(* IEC 61131-3 sources: daoli-st-library/DL_Algo (part 15) *)

(* ---- FB_DL_InputShaperZv.st ---- *)
(*
  ==================================================================
  组件名 Component  : FB_DL_InputShaperZv
  分类   Category   : DL_Algo
  复杂度 Complexity  : 中
  版本   Version    : 1.0.1
  功能   Purpose    : ZV（Zero Vibration）双脉冲输入整形器。按阻尼比 ζ 与固有频率
                      ωn 合成两脉冲序列（幅值 1/(1+A) 与 A/(1+A)，间隔 Δt），
                      触发沿到达时先出首脉冲，经 Δt 后出次脉冲，用于抑制指令
                      阶跃激起的残余振动。
  来源   Source     : self-std（公开控制理论 ZV 整形器语义）
  溯源   Origin     : ZV 输入整形属公开控制理论（Singer & Seering 公开文献语义），
                      道莅 clean-room 自研实现，未复制任何厂商私有库源码。
  平台   Platform   : 纯 IEC 61131-3（EXPT / SQRT / TON / R_TRIG / 标准转换函数）
  分工声明 Split     : 与 FB_DL_NotchFilter（反馈侧频域抑制属主）分工——后者对
                      测量信号做在线滤波；本件只整形前馈指令时序，不接管反馈、
                      不做滤波、不判机械到位。
  作者   Author     : 道莅代码库 · PLC 编程专家（R60）
  归属 Ownership     : E_DL_ZvPhase 属主为本文件（全库唯一定义，R264）；
                      引用件只引用不重声明（D13 返修补行）。
  ------------------------------------------------------------------
  边界 Boundary     :
                      一 时间口径单一化（R342）：Δt 内部一律以秒计算，转 TIME 时
                         统一乘 1000 后经 LREAL_TO_TIME 落毫秒，禁跨日历类型链；
                      二 采样约定：首脉冲在触发沿当拍输出，次脉冲在 Δt 到期拍
                         输出，两脉冲均为单拍（统一出口段每拍先预置 FALSE，R256）；
                      三 有限性闸显式枚举全部浮点输入（R272 自证：声明区 LREAL
                         输入共 2 个——fWn 与 fZeta——闸内逐个引用，无遗漏）；
                      四 域闸：fWn ≤ 0 判故障级码并冻结输出；ζ 域 [0, 0.95) 钳位，
                         越域置信息级码（ζ = 0 为无阻尼极限，取 A = 1 双等幅脉冲，
                         √(1−ζ²) = 1 结构性安全）；
                      五 使能 bEnable = FALSE 时语义为「冻结保持 + 清未决次脉冲」
                         （不再出脉冲，幅值与间隔保持末次有效值）——R191 声明行；
                      六 故障解除路径：eFault 相由复位沿迁回空闲并清锁存（bReset
                         为输入引脚，恒可达，R152 自证）；
                      七 时序滞后声明（D12 返修登记）：tonGap 的 PT 取上拍
                         _tDelay（段 0 刷新先于段 3 参数换算），ωn 突变拍 Δt
                         生效滞后一扫描拍；上层如需同拍生效，须在触发前一拍
                         稳定参数（显式声明，非遗漏）。
  错误码   Codes    :
    16#0002_0610【信息级】阻尼比 ζ 越域已钳位到 [0, 0.95)
    16#0002_0611【故障级】浮点入参非有限（NaN / Inf），输出冻结
    16#0002_0612【故障级】固有频率 ωn ≤ 0（域非法），输出冻结
  验收   Acceptance :
    算法已证（脚本）：未跑 ｜ 编译器已证（三平台）：未跑
    V1 ωn=10 rad/s、ζ=0 → A=1、幅值各 0.5、Δt=0.314159 s（314 ms）
    V2 ωn=10 rad/s、ζ=0.3 → A=0.371、幅值 0.7290/0.2710、Δt=0.3296 s
    V3 ζ=1.5 → 钳到 0.95、码 0610、序列仍出（bValid = TRUE）
    V4 ωn=0 → 码 0612、两脉冲恒假、eState = eFault
  修订记录 Revision  :
    2026-11-21  v1.0.0  R60 首版（批 2 · 序号 8）
    2026-11-21  v1.0.1  R61 返修：D12 边界段声明 tonGap PT 一拍滞后口径；
                        D13 补 E_DL_ZvPhase 属主 Ownership 行
  ==================================================================
*)

TYPE E_DL_ZvPhase :
(
    eIdle  := 0,  // 空闲：无未决次脉冲 / idle, no pending second pulse
    eWaitB := 10, // 等次脉冲：首脉冲已出，Δt 计时中 / waiting for the second pulse while the gap runs
    eFault := 20  // 故障：参数非法，输出冻结 / fault, the parameters are illegal and the outlet is frozen
);
END_TYPE

FUNCTION_BLOCK FB_DL_InputShaperZv
VAR_INPUT
    bEnable : BOOL := TRUE;       // 使能，FALSE 时冻结保持并清未决脉冲（边界五）/ the enable, false freezes and clears the pending pulse
    bTrig   : BOOL := FALSE;      // 整形触发电平，上升沿发起双脉冲序列 / the shaping trigger, the rising edge starts the pair
    bReset  : BOOL := FALSE;      // 复位沿：清故障锁存与未决序列并回空闲 / the reset edge, clears the latch and the pending pair
    fWn     : LREAL := 10.0;      // 固有角频率 [弧度每秒]，必须 > 0 / the natural angular frequency, must be positive
    fZeta   : LREAL := 0.1;       // 阻尼比 [-]，域 [0, 0.95) / the damping ratio inside the half open domain
END_VAR
VAR_OUTPUT
    bPulseA : BOOL := FALSE;      // 首脉冲单拍（触发沿当拍）[-] / the first pulse on the trigger scan
    bPulseB : BOOL := FALSE;      // 次脉冲单拍（Δt 到期拍）[-] / the second pulse on the expiry scan
    fAmpA   : LREAL := 0.5;       // 首脉冲幅值系数 [-]，与次脉冲之和为一 / the first amplitude coefficient
    fAmpB   : LREAL := 0.5;       // 次脉冲幅值系数 [-] / the second amplitude coefficient
    tDelay  : TIME := T#0S;       // 双脉冲间隔 Δt [毫秒] / the gap between the two pulses
    eState  : E_DL_ZvPhase;       // 主状态机当前态 [状态] / the current state of the main machine
    bValid  : BOOL := FALSE;      // 参数有效且序列可用标志 [-] / the parameters valid and the pair usable flag
    bError  : BOOL := FALSE;      // 故障锁存位 [-] / the latched fault bit
    eErr    : UDINT := 16#0000_0000; // 错误码，0 = 正常 / the error code, zero is ok
END_VAR
VAR
    _bInit    : BOOL := FALSE;                       // 首拍初始化标志（R310）/ the first scan flag
    _eState   : E_DL_ZvPhase := E_DL_ZvPhase.eIdle;  // 内部状态寄存器，段 4 唯一写点 / the internal state register, single writer
    _bPulseA  : BOOL := FALSE;                       // 首脉冲内部位，段 1 预清段 6 映射 / the internal first pulse bit, preset then mapped
    _bPulseB  : BOOL := FALSE;                       // 次脉冲内部位，段 1 预清段 6 映射 / the internal second pulse bit, preset then mapped
    _bPending : BOOL := FALSE;                       // 未决次脉冲位（间隔计时使能源）/ the pending second pulse flag driving the gap timer
    _bFault   : BOOL := FALSE;                       // 故障锁存副本（仅复位沿清除）/ the fault latch copy, cleared only on the reset edge
    _bFin     : BOOL := FALSE;                       // 浮点有限性闸结果（逐拍重算）/ the finiteness gate result, recomputed every scan
    _fZetaUse : LREAL := 0.0;                        // 钳位后的阻尼比工作副本 [-] / the clamped damping ratio copy
    _fA        : LREAL := 0.0;                       // 幅值比 A = exp(−ζπ/√(1−ζ²)) [-] / the amplitude ratio
    _fRoot     : LREAL := 1.0;                       // √(1−ζ²) 工作副本 [-] / the root working copy
    _fDtSec    : LREAL := 0.0;                       // 双脉冲间隔 [秒] / the gap in seconds
    _tDelay    : TIME := T#0S;                       // 内部间隔副本，段 6 单点映射 / the internal gap copy, mapped once in segment six
    rtTrig     : R_TRIG;                            // 触发沿实例，段 0 无条件刷新 / the trigger edge instance, refreshed unconditionally
    tonGap     : TON;                               // 间隔定时器，段 0 无条件刷新 / the gap timer, refreshed unconditionally
END_VAR
VAR CONSTANT
    DL_ZV_ZETAMAX : LREAL := 0.95;                  // 阻尼比上界（开区间）[-] / the damping ratio upper bound, exclusive
    DL_ZV_PI      : LREAL := 3.14159265358979323846; // 圆周率（LREAL 精度字面量，R51）/ the pi constant at the long real precision
    DL_ZV_E       : LREAL := 2.71828182845904523536; // 自然常数（EXPT 底数，禁厂商 EXP 方言）/ the natural base used with the standard power operator
    DL_ZV_MS      : LREAL := 1000.0;                // 秒到毫秒的换算因子 [毫秒每秒] / the seconds to milliseconds factor
END_VAR

// 段 0｜沿检测与间隔定时器无条件周期刷新（禁入分支，R7；IN 串故障锁存门控，FB50-1）/ segment 0, the unconditional refresh with the latch gate
rtTrig(CLK := bTrig); // 触发沿 / the trigger edge
tonGap(IN := _bPending AND _bFin AND (NOT _bFault), PT := _tDelay); // 间隔计时：未决且参数有效且无锁存 / the gap timing only while pending and valid

// 段 1｜首拍初始化与单拍标志预清（仅单拍标志入清单，R32 FB32-1；R256）/ segment 1, the first scan init and the one shot preset
IF NOT _bInit THEN // 首拍一拍 / the first scan
    _bInit := TRUE; // 置首拍标志 / raise the first scan flag
    _bPending := FALSE; // 未决位显式清零 / clear the pending flag explicitly
    _bFault := FALSE; // 故障锁存显式清零 / clear the fault latch explicitly
    _eState := E_DL_ZvPhase.eIdle; // 状态显式落空闲 / place the state to idle explicitly
END_IF
_bPulseA := FALSE; // 首脉冲预清零 / preset the first pulse false
_bPulseB := FALSE; // 次脉冲预清零 / preset the second pulse false

// 段 2｜参数有限性闸：显式枚举全部浮点输入 fWn 与 fZeta（R272 覆盖自证，边界三）/ segment 2, the finiteness gate enumerating every floating input
_bFin := (fWn = fWn) AND ((fWn - fWn) = (fWn - fWn)) AND (fZeta = fZeta) AND ((fZeta - fZeta) = (fZeta - fZeta)); // NaN 自反判 + Inf 差值自减判，两输入逐项 / the NaN reflexive and Inf difference tests on both inputs

// 段 3｜参数域闸：频率正域与阻尼比钳位（域闸覆盖参与换算的每个引脚，边界四）/ segment 3, the domain gate covering every pin used in the computation
IF NOT _bFin THEN // 非有限参数 / a non finite parameter
    _bFault := TRUE; // 锁存故障（段 5 迁移相）/ latch the fault, the segment five migrates the phase
ELSIF fWn <= 0.0 THEN // 频率域非法 / an illegal frequency domain
    _bFault := TRUE; // 锁存故障 / latch the fault
ELSE // 参数域合法：计算整形系数 / the parameters are legal, compute the shaping coefficients
    IF fZeta < 0.0 THEN // 阻尼比低于下界 / the damping below the floor
        _fZetaUse := 0.0; // 钳到零（无阻尼极限）/ clamp to zero, the undamped limit
    ELSIF fZeta >= DL_ZV_ZETAMAX THEN // 阻尼比达上界 / the damping at the bound
        _fZetaUse := 0.84375; // 钳到域几何内点 27/32（落在 [0, 0.95) 内，二级回退，R117）/ clamp to the interior point 27 over 32
    ELSE // 域内 / inside the domain
        _fZetaUse := fZeta; // 原值接管 / take the value as is
    END_IF
    _fRoot := SQRT(1.0 - _fZetaUse * _fZetaUse); // √(1−ζ²)：ζ ≤ 0.95 保证 > 0.31（结构性安全）/ the root is provably positive
    _fA := EXPT(DL_ZV_E, 0.0 - _fZetaUse * DL_ZV_PI / _fRoot); // A = exp(−ζπ/√(1−ζ²)) / the amplitude ratio
    fAmpA := 1.0 / (1.0 + _fA); // 首脉冲幅值（除子 ≥ 1 恒正）/ the first coefficient with a divisor of at least one
    fAmpB := _fA / (1.0 + _fA); // 次脉冲幅值 / the second coefficient
    _fDtSec := DL_ZV_PI / (fWn * _fRoot); // Δt = π/(ωn√(1−ζ²)) [秒] / the gap in seconds
    _tDelay := LREAL_TO_TIME(_fDtSec * DL_ZV_MS); // 秒口径单一化后落毫秒（R342）/ the single second domain converted to milliseconds
END_IF

// 段 4｜主状态机（ENUM + CASE，ELSE 拦非法态）/ segment 4, the main machine with the illegal state guard
CASE _eState OF
    E_DL_ZvPhase.eIdle: // 空闲相：等触发沿 / the idle phase waiting for the trigger edge
        IF bEnable AND _bFin AND (NOT _bFault) AND (fWn > 0.0) AND rtTrig.Q THEN // 迁入判据带全量闸位复检（R274）/ the entry with the full gate recheck
            _bPulseA := TRUE; // 首脉冲（触发沿当拍，边界二）/ the first pulse on the trigger scan
            _bPending := TRUE; // 置未决次脉冲 / raise the pending second pulse
            _eState := E_DL_ZvPhase.eWaitB; // 迁入等次脉冲相 / enter the waiting phase
        END_IF
    E_DL_ZvPhase.eWaitB: // 等次脉冲相 / the waiting phase
        IF tonGap.Q THEN // 间隔到期：出次脉冲 / the gap expired, raise the second pulse
            _bPulseB := TRUE; // 次脉冲单拍 / the second pulse
            _bPending := FALSE; // 清未决位 / clear the pending flag
            _eState := E_DL_ZvPhase.eIdle; // 迁回空闲 / back to idle
        ELSIF (NOT bEnable) OR (NOT _bFin) OR _bFault THEN // 出口二：失能 / 参数转非有限 / 锁存（前置条件消失）/ the second exit with the prerequisite gone
            _bPending := FALSE; // 清未决位（弃用序列，不出次脉冲）/ discard the pending pair
            _eState := E_DL_ZvPhase.eIdle; // 迁回空闲 / back to idle
        END_IF
    E_DL_ZvPhase.eFault: // 故障相：锁存保持，等复位沿（解除可达，边界六）/ the fault phase held until the reset edge
        IF bReset THEN // 复位电平（复位作用域：清锁存 + 清未决 + 迁相位）/ the reset with the declared scope
            _bFault := FALSE; // 清故障锁存 / clear the fault latch
            _bPending := FALSE; // 清未决序列 / clear the pending pair
            _eState := E_DL_ZvPhase.eIdle; // 故障相迁出边回空闲 / the exit edge back to idle
        END_IF
    ELSE // 非法枚举值拦截 / the illegal enumeration guard
        _eState := E_DL_ZvPhase.eIdle; // 落回空闲 / force back to idle
        _bFault := TRUE; // 置故障锁存 / latch the fault
END_CASE

// 段 5｜故障锁存迁移闸（置于解除段之后防同拍抢迁，R258）/ segment 5, the fault latch to phase gate placed after the release
IF _bFault AND (_eState <> E_DL_ZvPhase.eFault) THEN // 已锁存但不在故障相 / latched but not in the fault phase
    _eState := E_DL_ZvPhase.eFault; // 迁入故障相 / enter the fault phase
END_IF

// 段 6｜统一出口（内部副本单点映射，R180；故障码锁存回放，R187）/ segment 6, the unified outlet
bPulseA := _bPulseA AND bEnable; // 首脉冲出口（失能不出脉冲）/ the first pulse outlet gated by the enable
bPulseB := _bPulseB AND bEnable; // 次脉冲出口（失能不出脉冲）/ the second pulse outlet gated by the enable
tDelay := _tDelay; // 间隔出口 / the gap outlet
eState := _eState; // 状态出口 / the state outlet
bError := _bFault; // 故障位出口（与锁存同源）/ the fault bit outlet from the same latch
bValid := _bFin AND (fWn > 0.0) AND (NOT _bFault); // 参数可用标志（逐拍重算）/ the usable flag recomputed every scan
IF _bFault THEN // 故障锁存回放优先 / the latched fault replays first
    IF NOT _bFin THEN // 非有限成因（独立码值，R190）/ the non finite cause with its own code
        eErr := 16#0002_0611; // 故障级：浮点入参非有限 / fault grade, a non finite floating input
    ELSE // 频率域成因 / the frequency domain cause
        eErr := 16#0002_0612; // 故障级：固有频率非正 / fault grade, the natural frequency is not positive
    END_IF
ELSIF ABS(_fZetaUse - fZeta) > 1.0E-9 THEN // 阻尼比被钳位（浮点差值比较，禁等号；信息级逐拍重算）/ the damping clamped, compared by tolerance
    eErr := 16#0002_0610; // 信息级：阻尼比越域已钳位 / informational, the damping clamped
    bError := FALSE; // 信息级不置 bError（R45 配对口径：仅故障级置位）/ the informational code never raises the fault bit
ELSE // 无事件 / no event
    eErr := 16#0000_0000; // 正常 / ok
END_IF
END_FUNCTION_BLOCK

(* ---- FB_DL_Integrator.st ---- *)
(*==============================================================================
 * 组件名称 (Component)  : FB_DL_Integrator
 * 所属子库 (Sublibrary) : DL_Algo
 * 当前版本 (Version)    : 1.0.1
 * 兼容性   (Platform)   : CODESYS 3.5 / TwinCAT 3 / 汇川 InoProShop / Machine Expert
 *                         仅依赖 Standard.library（MIN / MAX / ABS / LREAL_TO_REAL），零厂商方言
 * 功能描述 (Function)   : 梯形法离散积分器：fSum += (fIn + fInPrev)/2 · fDt，
 *                         精度高于矩形法，对缓变信号无系统偏差。内部以 LREAL
 *                         双精度累加、输出转 REAL，防长时累计的舍入漂移。
 *                         带上下限限幅（触限保持）、保持（bHold）、电平复位
 *                         （bReset）、跟踪回投（bTrack）。现场用途：流量累计
 *                         （总量表）、速度→位移、电量/电能累计。
 * 开源溯源 (Origin)     : 原创实现。双精度累加思想源自 OSCAT Basic 的
 *                         FT_INT2 误差抑制行为定义（EPL-2.0），clean-room
 *                         编写，未复制任何源码。
 * 本文件内含       : TYPE  E_DL_IntState（配套枚举，归属 DL_Algo）
 *                    FB    FB_DL_Integrator
 * 依赖     (Depends)    : 无 DL_ 内部依赖；Standard.library: LREAL_TO_REAL
 * 红线自检 (Redline)    : R1 ✓ 零全局变量表与外部变量引用 ｜ R2 ✓ 零物理 IO 地址直写
 *                         R3 ✓ 纯 IEC 61131-3 ｜ R4 ✓ 量程对调+溢出钳位+非有限值拒绝
 *                         R5 ✓ 全变量中英双语同行注释 ｜ R6 ✓ 五态 ENUM+CASE+ELSE
 *                         R7 N/A（无定时器/边沿实例）
 * 【边界披露 / Boundary disclosure】
 *   B1 rOutMin > rOutMax：自动对调并置 16#0002_0001，不中断扫描。
 *   B2 复位优先于积分：bReset 电平触发，复位拍不积分（先判 bReset）。
 *   B3 输入非有限值（NaN 或幅值超 1.0E30）：本拍拒绝积分、保持累加器、
 *      fInPrev 不同步，置 16#0002_0004。
 *   B4 累加器幅值超 1.0E30：强制钳位防 LREAL 溢出，置 16#0002_0001。
 *   B5 保持期（bHold 或未使能）不积分，fInPrev 亦不更新，恢复时无历史跳变。
 *   B6 触限后每拍仍尝试积分：输入反向或限幅放宽时自动恢复，无需复位。
 * 【验收向量 / Acceptance vectors】
 *   V1  fIn=10 EU 恒定，tSampleTime=100MS，1s 后 fOut≈10 EU·s（梯形法与
 *       解析值一致，矩形法会偏 0.5 EU·s，对比可见梯形优势）
 *   V2  fIn 由 0 线性升至 10（每拍 +1），1s 后 fOut≈5.05 EU·s（与解析积分一致）
 *   V3  rOutMax=3，V1 持续 → fOut 钳位 3、bLimitHigh=TRUE、状态 eLimited
 *   V4  bHold=TRUE → fOut 冻结；释放后从冻结值继续
 *   V5  bReset 一拍 → fOut=0、fInPrev 同步当前输入（防复位后首拍尖峰）
 *   V6  bTrack 一拍（fTrackValue=100）→ fOut=100，无扰动回投
 *   V7  fIn=NaN → 16#0002_0004，fOut 保持，累加器不动
 * 修订历史 (Revision)   :
 *   2026-11-15  v1.0.0  首版入库（Round 04 · Phase 3 · DL_Algo 批次）
 *   2026-11-15  v1.0.1  阶段五终审精修：首扫自动跟踪判据修复（原 bInit 判据
 *                       反向，bTrack 一次后累加器被永久锁死为跟踪值）
 *============================================================================*)

(*-----------------------------------------------------------------------------
 * 枚举: E_DL_IntState（归属 DL_Algo，与 FB_DL_Integrator 同文件）
 * 含义: 积分器状态机离散状态。数值步长留空位便于后续插态而不破坏已有工程。
 *----------------------------------------------------------------------------*)
TYPE E_DL_IntState :
(
    eIdle        := 0,   // 空闲态：未使能，累加器保持 / Idle state, accumulator held
    eHold        := 10,  // 保持态：操作员请求冻结累加 / Hold state, accumulation frozen on request
    eIntegrating := 20,  // 积分态：梯形法逐拍累加 / Integrating, trapezoidal accumulation
    eLimited     := 30,  // 触限态：累加器停在限幅值，反向输入自动恢复 / Limited, auto recovers on reverse input
    eFault       := 99   // 故障兜底态：非法状态拦截，自动回空闲 / Fault fallback, auto recover to idle
);
END_TYPE

(*==============================================================================
 * 功能块: FB_DL_Integrator
 * 调用约定: 每个扫描周期无条件调用一次；bReset 电平触发（保持 TRUE 即持续清零）。
 * 无状态泄漏: 全部状态驻留于实例私有 VAR，可多实例并行互不影响。
 * 精度披露: 内部 LREAL 双精度累加、每拍输出转 REAL；单位为 [EU·s]
 *           （被积量 [EU] × 时间 [s]），总表类应用注意换算口径。
 *============================================================================*)
FUNCTION_BLOCK FB_DL_Integrator
VAR_INPUT
    bEnable     : BOOL := FALSE;      // 使能标志，FALSE 保持累加器 / Enable flag, FALSE holds accumulator
    fIn         : REAL := 0.0;        // 被积量 [EU]，如流量/速度/电流 / Integrated input [EU]
    rOutMin     : REAL := 0.0;        // 积分下限 [EU·s]，大于上限时自动对调 / Integral lower limit [EU·s], swapped if greater
    rOutMax     : REAL := 1.0E12;     // 积分上限 [EU·s]，长时累计防溢出 / Integral upper limit [EU·s]
    bHold       : BOOL := FALSE;      // 保持请求，TRUE 冻结累加 / Hold request, TRUE freezes accumulation
    bReset      : BOOL := FALSE;      // 复位信号，电平触发清零 / Reset signal, level triggered clear
    bTrack      : BOOL := FALSE;      // 跟踪使能，TRUE 时累加器立即跟随 fTrackValue / Track enable, accumulator follows track value
    fTrackValue : REAL := 0.0;        // 跟踪值 [EU·s]，投切无扰动基准 / Track value [EU·s], bumpless transfer reference
    tSampleTime : TIME := T#100MS;    // 采样周期 [s]，小于 10ms 钳位为 10ms / Sample time [s], clamped to 10ms
END_VAR
VAR_OUTPUT
    fOut        : REAL;               // 积分结果 [EU·s] / Integration result [EU·s]
    bLimitHigh  : BOOL;               // 触上限标志 / Upper limit reached flag
    bLimitLow   : BOOL;               // 触下限标志 / Lower limit reached flag
    bError      : BOOL;               // 故障标志（瞬时，逐拍重算） / Fault flag, transient, recomputed every scan
    uErrorId    : UDINT;              // 故障码，0 = 无故障 / Error code, 0 = no error
END_VAR
VAR
    fSumLReal   : LREAL;              // 双精度累加器 [EU·s] / Double precision accumulator [EU·s]
    fInPrev     : REAL;               // 上一拍被积量 [EU]，梯形法端点 / Previous input [EU], trapezoid endpoint
    fDt         : REAL;               // 折算后的采样周期 [s] / Converted sample period [s]
    bInFinite   : BOOL;               // 本拍输入有限值标志 / Input finite validity flag this scan
    bInit       : BOOL;               // 首扫标志：首扫自动跟踪 / First scan flag, auto track on first scan
    eState      : E_DL_IntState;      // 主状态机当前状态 / Current state of the main state machine
END_VAR
VAR CONSTANT
    DL_INT_ABS_MAX : LREAL := 1.0E30; // 累加器幅值上限 [EU·s]，防溢出 / Accumulator magnitude limit [EU·s]
END_VAR

(*------------------------------------------------------------------------------
 * 段 1｜公共参数处理（通用约定 0-1/0-2）：周期钳位、量程对调、故障码瞬时清零
 *      Common handling: sample time clamp, limit swap, transient code reset
 *-----------------------------------------------------------------------------*)
uErrorId   := 16#0000_0000;         // 故障码逐拍重算 / Error code recomputed every scan
bError     := FALSE;                // 故障标志逐拍重算 / Fault flag recomputed every scan
bLimitHigh := FALSE;                // 触限标志逐拍重算 / Limit flags recomputed every scan
bLimitLow  := FALSE;                // 触限标志逐拍重算 / Limit flags recomputed every scan

IF tSampleTime < T#10MS THEN
    fDt      := TIME_TO_REAL(T#10MS) / 1000.0; // 非法周期钳位为 10ms / Illegal period clamped to 10ms
    uErrorId := 16#0002_0002;           // 采样周期非法已钳位 / Sample time illegal, clamped
ELSE
    fDt      := TIME_TO_REAL(tSampleTime) / 1000.0; // 周期换算为秒 [s] / Period converted to seconds [s]
END_IF

IF rOutMin > rOutMax THEN
    rOutMin   := rOutMin + rOutMax;     // 三步对调第一步：求和 / Swap step one: sum
    rOutMax   := rOutMin - rOutMax;     // 三步对调第二步：得旧下限 / Swap step two: old lower limit
    rOutMin   := rOutMin - rOutMax;     // 三步对调第三步：得旧上限 / Swap step three: old upper limit
    uErrorId  := 16#0002_0001;          // 参数越界已对调 / Limits out of order, swapped
END_IF

(*------------------------------------------------------------------------------
 * 段 2｜输入合法性与复位/跟踪（边界 B2/B3、约定 0-6）
 *      Input validity and reset/track handling
 *-----------------------------------------------------------------------------*)
bInFinite := NOT (fIn <> fIn) AND (ABS(fIn) <= 1.0E30); // NaN 判别 + 幅值防御 / NaN check plus magnitude guard

IF NOT bInFinite THEN
    uErrorId := 16#0002_0004;           // 输入非有限值已拒绝 / Non-finite input rejected
END_IF

IF bTrack OR (NOT bInit) THEN
    fSumLReal := MIN(MAX(fTrackValue, rOutMin), rOutMax); // 累加器立即跟随跟踪值并限幅 / Accumulator follows track value with limits
    IF bInFinite THEN
        fInPrev := fIn;                 // 端点同步当前输入 / Endpoint synced to current input
    END_IF
    eState := eIdle;                    // 回空闲重新评估 / Back to idle for re-evaluation
    bInit  := TRUE;                     // 首扫标志置位 / First scan flag set
END_IF

IF bReset THEN
    fSumLReal := 0.0;                   // 复位优先：累加器清零 / Reset priority: accumulator cleared
    IF bInFinite THEN
        fInPrev := fIn;                 // 端点同步当前输入，防复位后尖峰 / Endpoint synced, prevents post-reset spike
    END_IF
    eState := eIdle;                    // 复位后回空闲 / Back to idle after reset
END_IF

IF NOT bEnable THEN
    eState := eIdle;                    // 未使能：强制空闲、累加器保持 / Disabled: force idle, accumulator held
END_IF

(*------------------------------------------------------------------------------
 * 段 3｜主状态机（红线 R6）：五态 ENUM + CASE + ELSE 兜底
 *      Main state machine: five-state ENUM + CASE with mandatory ELSE fallback
 *-----------------------------------------------------------------------------*)
CASE eState OF

    eIdle:  // 空闲态：使能且输入有效且未复位未保持 → 进入积分态 / Idle: enter integrating when conditions met
        IF bEnable AND bInFinite AND (NOT bReset) AND (NOT bHold) THEN
            eState := eIntegrating;     // 进入积分态（本拍先迁移，下拍起积分）/ Enter integrating, integrate from next scan
        END_IF

    eHold:  // 保持态：释放后回积分态 / Hold: resume integrating after release
        IF bEnable AND bInFinite AND (NOT bReset) AND (NOT bHold) THEN
            eState := eIntegrating;     // 恢复积分 / Resume integration
        ELSIF NOT bEnable THEN
            eState := eIdle;            // 使能跌落回空闲 / Back to idle when disabled
        END_IF

    eIntegrating:  // 积分态：梯形法逐拍累加（边界 B3 拒绝非有限值）/ Integrating: trapezoidal accumulation
        IF NOT bEnable THEN
            eState := eIdle;            // 使能跌落回空闲 / Back to idle when disabled
        ELSIF bHold THEN
            eState := eHold;            // 保持请求 / Hold request
        ELSIF bInFinite THEN
            fSumLReal := fSumLReal + (fIn + fInPrev) / 2.0 * fDt; // 梯形法累加 [EU·s] / Trapezoidal accumulation [EU·s]
            fInPrev    := fIn;          // 端点更新 / Endpoint updated
        END_IF

    eLimited:  // 触限态：每拍仍尝试积分，反向输入或限幅放宽时自动恢复（边界 B6）/ Limited: retry every scan, auto recover
        IF NOT bEnable THEN
            eState := eIdle;            // 使能跌落回空闲 / Back to idle when disabled
        ELSIF bHold THEN
            eState := eHold;            // 保持请求 / Hold request
        ELSIF bInFinite THEN
            fSumLReal := fSumLReal + (fIn + fInPrev) / 2.0 * fDt; // 继续累加（限幅兜底）/ Keep accumulating, clamp guards
            fInPrev    := fIn;          // 端点更新 / Endpoint updated
        END_IF

    eFault:  // 故障兜底态：累加器保持，自动回空闲（无锁死）/ Fault fallback: accumulator held, recover to idle
        eState := eIdle;                // 自动恢复空闲 / Auto recover to idle

    ELSE  // 非法状态拦截：任何未定义状态一律进故障态并置码 / Illegal state interception
        eState   := eFault;             // 强制故障态 / Force fault state
        uErrorId := 16#0002_0005;       // 非法状态兜底 / Illegal state fallback
        bError   := TRUE;               // 故障标志置位 / Fault flag set

END_CASE;

(*------------------------------------------------------------------------------
 * 段 4｜溢出钳位与量程限幅、输出整形（边界 B4/B1）
 *      Overflow clamp, range limiting and output shaping
 *-----------------------------------------------------------------------------*)
IF fSumLReal > DL_INT_ABS_MAX THEN
    fSumLReal := DL_INT_ABS_MAX;        // 幅值超限钳位防溢出 / Magnitude clamped against overflow
    uErrorId  := 16#0002_0001;          // 参数越界已钳位 / Value out of range, clamped
END_IF
IF fSumLReal < -DL_INT_ABS_MAX THEN
    fSumLReal := -DL_INT_ABS_MAX;       // 负向幅值钳位 / Negative magnitude clamped
    uErrorId  := 16#0002_0001;          // 参数越界已钳位 / Value out of range, clamped
END_IF

IF fSumLReal >= rOutMax THEN
    fSumLReal   := rOutMax;             // 触上限钳位 / Clamped at upper limit
    bLimitHigh  := TRUE;                // 触上限标志 / Upper limit flag
    IF bEnable AND (NOT bHold) THEN
        eState := eLimited;             // 进入触限态 / Enter limited state
    END_IF
END_IF
IF fSumLReal <= rOutMin THEN
    fSumLReal  := rOutMin;              // 触下限钳位 / Clamped at lower limit
    bLimitLow  := TRUE;                 // 触下限标志 / Lower limit flag
    IF bEnable AND (NOT bHold) THEN
        eState := eLimited;             // 进入触限态 / Enter limited state
    END_IF
END_IF

fOut := LREAL_TO_REAL(fSumLReal);       // 双精度累加器转 REAL 输出 [EU·s] / Accumulator converted to REAL output [EU·s]
END_FUNCTION_BLOCK

(* ---- FB_DL_IterSolverRunner.st ---- *)
(* ============================================================
   DL_Algo / FB_DL_IterSolverRunner ｜ v1.0.0 ｜ 2026-11-25
   功能：多方法求根运行器（0 二分 / 1 试位 / 2 割线 / 3 Illinois / 4 Brent）
         ＋括号管理＋无解与超时出口＋迭代上限防死锁。
         纯 IEC 无函数指针，采用「求值回灌协议」：本件在 fXOut 给出待求值点，
         调用方求残差后调用方法 FeedEval(fX, fF) 回灌，主体下一拍消费并给下一点。
   边界：① 括号两端同号 → eFail、码 5（无解），不空转；② 迭代上限（0=不限，默认 100）与
         总超时（0=不限，默认 T#5S）双防死锁，各自独立码（R190 归因唯一）；超时狗武装域
         覆盖 eEvalLo / eEvalHi / eRun 三相，求值相回灌断链亦能超时退出，不永久挂死；
         ③ 回灌点与待求值点
         不匹配（|Δx|>1E-9）→ 丢弃不置错；④ 复位沿作用域：清括号/计数/回灌位/锁存/
         相位，不动 _bInit；⑤ 出口非有限即落 0（N1）；⑥ 方法内不驻留跨拍状态。
   依赖：仅 IEC 61131-3（TON/R_TRIG/ABS/MIN/MAX/LIMIT）
   溯源：DLF-B-ROOTSTEP（内部原创线）｜枚举归属：E_DL_IterRunnerPhase 唯一属主
   码位：零 16# 范式；uErrId 0 无 / 1 组态 / 2 非有限 / 3 迭代上限 / 4 超时 /
         5 括号同号 / 6 非法相位
   ============================================================ *)
TYPE E_DL_IterRunnerPhase :
(
    eIdle   := 0,    // 待机：等待启动沿 / Idle, waiting for the start edge
    eEvalLo := 10,   // 求值下界：等 f(xLo) 回灌 / Waiting for the lower bound residual
    eEvalHi := 20,   // 求值上界：等 f(xHi) 回灌 / Waiting for the upper bound residual
    eRun    := 30,   // 迭代：给试算点并消费回灌 / Iterating over trial points
    eDone   := 40,   // 完成：宽度或残差达标 / Finished within tolerance
    eFail   := 50,   // 失败：无解 / 上限 / 超时 / Failed by no root, cap or timeout
    eFault  := 90    // 故障：组态或非有限锁存 / Fault latched
);
END_TYPE

FUNCTION_BLOCK FB_DL_IterSolverRunner
VAR_INPUT
    bStart   : BOOL;   // 启动，上升沿开始一轮 [-] / Start on the rising edge
    bReset   : BOOL;   // 复位，上升沿解除失败与故障 [-] / Reset on the rising edge
    fXLo     : LREAL;  // 初始括号下界 [-] / Initial lower bracket bound
    fXHi     : LREAL;  // 初始括号上界 [-] / Initial upper bracket bound
    fTol     : LREAL;  // 宽度收敛容差，域 > 0 [-] / Convergence tolerance on the width
    nMethod  : INT;    // 方法选择 0..4 [-] / Method selector
    nIterMax : INT := 100;         // 迭代上限，0 = 不限，默认 100 次（防死锁）[次] / Iteration cap, zero means unlimited
    tTimeout : TIME := T#5S;       // 总超时，0 = 不限，默认 5s（防死锁）[ms] / Overall timeout, zero means unlimited
END_VAR
VAR_OUTPUT
    bDone    : BOOL;   // 求根完成 [-] / Root finding finished
    bError   : BOOL;   // 失败或故障 [-] / Failed or faulted
    fXOut    : LREAL;  // 当前待求值点（完成时为根候选）[-] / Point to evaluate
    fResid   : LREAL;  // 末次回灌残差 [-] / Last residual fed back
    uErrId   : UDINT;  // 事件码，0 = 无事件 [-] / Event code
    nIterOut : INT;    // 已用迭代次数 [次] / Iterations consumed
END_VAR
VAR
    rtStart  : R_TRIG;                                           // 启动沿实例，段 0 无条件刷新 / Start edge
    rtReset  : R_TRIG;                                           // 复位沿实例，段 0 无条件刷新 / Reset edge
    tonTotal : TON;                                              // 总超时狗，段 0 无条件刷新 / Overall watchdog
    _eState  : E_DL_IterRunnerPhase := E_DL_IterRunnerPhase.eIdle; // 内部相位 / Internal phase
    _bInit   : BOOL := FALSE;                                    // 首扫初始化已执行 [-] / First scan init done
    _bFed    : BOOL := FALSE;                                    // 回灌到位（协议位，方法置位）[-] / Feedback ready
    _fFedX   : LREAL := 0.0;                                     // 回灌点横坐标 [-] / Fed back abscissa
    _fFedF   : LREAL := 0.0;                                     // 回灌残差 [-] / Fed back residual
    _fA      : LREAL := 0.0;                                     // 括号下界 [-] / Lower bracket bound
    _fB      : LREAL := 0.0;                                     // 括号上界 [-] / Upper bracket bound
    _fFa     : LREAL := 0.0;                                     // 下界残差 [-] / Residual at the lower bound
    _fFb     : LREAL := 0.0;                                     // 上界残差 [-] / Residual at the upper bound
    _fXCur   : LREAL := 0.0;                                     // 当前待求值点 [-] / Current point to evaluate
    _nIter   : INT := 0;                                         // 已用迭代次数 [次] / Iterations consumed
    _bFault  : BOOL := FALSE;                                    // 故障锁存位 [-] / Latched fault bit
    _bFail   : BOOL := FALSE;                                    // 失败锁存位 [-] / Latched failure bit
    _uFault  : UDINT := 0;                                       // 事件码锁存 [-] / Latched event code
    _bCfgBad : BOOL;                                             // 组态非法当拍量 [-] / Illegal configuration flag
    _bNonFin : BOOL;                                             // 入参非有限当拍量 [-] / Non-finite argument flag
    _bTmoArm : BOOL;                                             // 总超时狗武装量（三相驻留 TRUE）[-] / Watchdog arming flag
END_VAR
VAR CONSTANT
    DL_ISR_EPS : LREAL := 1.0E-9;  // 回灌点匹配与判零容差 [-] / Feedback match and zero tolerance
    DL_ISR_C_CFG : UDINT := 1;     // 码 1：组态非法 / Code one, illegal configuration
    DL_ISR_C_FIN : UDINT := 2;     // 码 2：非有限 / Code two, non-finite value
    DL_ISR_C_ITER : UDINT := 3;    // 码 3：迭代上限 / Code three, iteration cap reached
    DL_ISR_C_TMO : UDINT := 4;     // 码 4：总超时 / Code four, overall timeout
    DL_ISR_C_SGN : UDINT := 5;     // 码 5：括号同号 / Code five, bracket lost by equal signs
    DL_ISR_C_ILL : UDINT := 6;     // 码 6：非法相位 / Code six, illegal phase fallback
END_VAR

(* 方法 NextTrial：按方法选择给下一个试算点，回退固定为括号中点（必能推进）。
   参数全部经引脚传入，不访问 FB 成员，方法内无跨拍状态（R3 方法准则）。 *)
METHOD NextTrial : LREAL
VAR_INPUT
    nSel   : INT;    // 方法选择 0..4 [-] / Method selector
    fA     : LREAL;  // 括号下界 [-] / Lower bracket bound
    fB     : LREAL;  // 括号上界 [-] / Upper bracket bound
    fFa    : LREAL;  // 下界残差 [-] / Residual at the lower bound
    fFb    : LREAL;  // 上界残差 [-] / Residual at the upper bound
    fXPrev : LREAL;  // 上一步试算点 [-] / Previous trial point
    fFxPrev : LREAL; // 上一步残差 [-] / Residual at the previous trial point
END_VAR
VAR
    _fLo  : LREAL;  // 括号小端 [-] / Smaller bracket end
    _fHi  : LREAL;  // 括号大端 [-] / Larger bracket end
    _fMid : LREAL;  // 中点 [-] / Midpoint
    _fDen : LREAL;  // 差分分母 [-] / Slope denominator
    _fX   : LREAL;  // 试算点暂存 [-] / Staged trial point
END_VAR

_fLo := MIN(fA, fB);  _fHi := MAX(fA, fB);
_fMid := _fLo + (_fHi - _fLo) / 2.0;
_fX := _fMid;                                  // 缺省回退中点
CASE nSel OF
0:  _fX := _fMid;                              // 二分
1:  _fDen := fFb - fFa;                        // 试位
    IF ABS(_fDen) > DL_ISR_EPS THEN _fX := fA - fFa * (fB - fA) / _fDen; END_IF
2:  _fDen := fFxPrev - fFa;                    // 割线（最近两点差商）
    IF ABS(_fDen) > DL_ISR_EPS THEN _fX := fXPrev - fFxPrev * (fXPrev - fA) / _fDen; END_IF
3:  _fDen := (fFb / 2.0) - fFa;                // Illinois（停滞端折半）
    IF ABS(_fDen) > DL_ISR_EPS THEN _fX := fA - fFa * (fB - fA) / _fDen; END_IF
4:  IF (ABS(fFa - fFb) > DL_ISR_EPS) AND (ABS(fFa - fFxPrev) > DL_ISR_EPS)
       AND (ABS(fFb - fFxPrev) > DL_ISR_EPS) THEN   // Brent：逆二次插值
        _fX := fA * (fFb * fFxPrev) / ((fFa - fFb) * (fFa - fFxPrev))
             + fB * (fFa * fFxPrev) / ((fFb - fFa) * (fFb - fFxPrev))
             + fXPrev * (fFa * fFb) / ((fFxPrev - fFa) * (fFxPrev - fFb));
    END_IF
ELSE
    _fX := _fMid;                              // 非法方法号：回退二分
END_CASE
IF (_fX <> _fX) OR ((_fX - _fX) <> (_fX - _fX)) THEN
    NextTrial := _fMid;                        // 非有限：回退中点
ELSE
    NextTrial := LIMIT(_fLo, _fX, _fHi);       // 夹界即 N4 出口闸
END_IF
END_METHOD

(* 方法 FeedEval：调用方回灌残差。仅接受与本拍待求值点匹配的回灌（防陈旧值污染
   括号）；不匹配静默丢弃；本方法不推进相位（推进在主体 CASE）。 *)
METHOD FeedEval : BOOL
VAR_INPUT
    fX : LREAL;  // 求值点横坐标 [-] / Abscissa the host evaluated
    fF : LREAL;  // 该点残差 [-] / Residual at that abscissa
END_VAR

FeedEval := FALSE;
IF (fX <> fX) OR (fF <> fF) THEN RETURN; END_IF
IF ABS(fX - _fXCur) > DL_ISR_EPS THEN RETURN; END_IF
_fFedX := fX;  _fFedF := fF;  _bFed := TRUE;  FeedEval := TRUE;
END_METHOD

(* 段 0：沿实例与定时器无条件每拍刷新（R7） *)
rtStart (CLK := bStart);
rtReset (CLK := bReset);
(* 超时狗武装域 = 三相驻留（eEvalLo / eEvalHi / eRun）：只守 eRun 时求值相漏回灌即永久挂死无码 *)
_bTmoArm := (_eState = E_DL_IterRunnerPhase.eEvalLo)
            OR (_eState = E_DL_IterRunnerPhase.eEvalHi)
            OR (_eState = E_DL_IterRunnerPhase.eRun);
tonTotal (IN := _bTmoArm AND (NOT _bFault) AND (tTimeout > T#0S),
          PT := tTimeout);                     // tTimeout = 0 表示不限超时

(* 段 1：单拍量预清零（锁存量与回灌位不入清单，R107） *)
_bCfgBad := FALSE;  _bNonFin := FALSE;

(* 段 2：首扫与复位沿同款初始化（清锁存 / 清括号与计数 / 迁相位，R310/R311） *)
IF (NOT _bInit) OR rtReset.Q THEN
    _bInit := TRUE;  _bFault := FALSE;  _bFail := FALSE;  _uFault := 0;
    _bFed := FALSE;  _nIter := 0;  _fA := 0.0;  _fB := 0.0;  _fXCur := 0.0;
    _eState := E_DL_IterRunnerPhase.eIdle;
END_IF

(* 段 3：组态闸与非有限闸（覆盖全部参与判据的引脚，R272） *)
IF (fTol <= 0.0) OR (nMethod < 0) OR (nMethod > 4) OR (nIterMax < 0) THEN _bCfgBad := TRUE; END_IF
IF (fXLo <> fXLo) OR (fXHi <> fXHi) OR (fTol <> fTol) THEN _bNonFin := TRUE; END_IF
(* Inf 双判（正负无穷括号 = 组态非法，禁带入括号管理）：判据与出口同源于原始入参 *)
IF ((fXLo - fXLo) <> (fXLo - fXLo)) OR ((fXHi - fXHi) <> (fXHi - fXHi))
   OR ((fTol - fTol) <> (fTol - fTol)) THEN _bNonFin := TRUE; END_IF
IF (_bCfgBad OR _bNonFin) AND (NOT (_bFault OR _bFail)) THEN
    _bFault := TRUE;  _eState := E_DL_IterRunnerPhase.eFault;
    IF _bNonFin THEN
        _uFault := DL_ISR_C_FIN;      // 非有限优先归因（值与判据同源，N1）
    ELSE
        _uFault := DL_ISR_C_CFG;      // 组态非法：容差/方法号/迭代上限
    END_IF
END_IF

(* 段 4：主状态机（七相全覆盖 + ELSE 非法相位兜底） *)
CASE _eState OF

E_DL_IterRunnerPhase.eIdle:
    IF rtStart.Q THEN
        _fA := fXLo;  _fB := fXHi;  _nIter := 0;  _bFed := FALSE;
        _fXCur := fXLo;  _eState := E_DL_IterRunnerPhase.eEvalLo;   // 先求下界残差
    END_IF

E_DL_IterRunnerPhase.eEvalLo:
    IF _bFed THEN                              // 事件：回灌到位
        _fFa := _fFedF;  _bFed := FALSE;  _fXCur := _fB;
        _eState := E_DL_IterRunnerPhase.eEvalHi;
    ELSIF tonTotal.Q THEN                      // 事件缺失：超时接管（回灌断链不再永久挂死）
        _bFail := TRUE;  _uFault := DL_ISR_C_TMO;  _eState := E_DL_IterRunnerPhase.eFail;
    ELSIF ABS(_fB - _fA) <= DL_ISR_EPS THEN    // 前置消失：括号零宽
        _bFail := TRUE;  _uFault := DL_ISR_C_SGN;  _eState := E_DL_IterRunnerPhase.eFail;
    END_IF

E_DL_IterRunnerPhase.eEvalHi:
    IF _bFed THEN
        _fFb := _fFedF;  _bFed := FALSE;
        IF (ABS(_fFa) <= DL_ISR_EPS) OR (ABS(_fFb) <= DL_ISR_EPS) THEN
            _eState := E_DL_IterRunnerPhase.eDone;          // 端点已是根
        ELSIF ((_fFa > 0.0) AND (_fFb > 0.0)) OR ((_fFa < 0.0) AND (_fFb < 0.0)) THEN
            _bFail := TRUE;  _uFault := DL_ISR_C_SGN;       // 同号：无解归因
            _eState := E_DL_IterRunnerPhase.eFail;
        ELSE
            _fXCur := NextTrial(nSel := nMethod, fA := _fA, fB := _fB, fFa := _fFa,
                                fFb := _fFb, fXPrev := _fA, fFxPrev := _fFa);
            _eState := E_DL_IterRunnerPhase.eRun;
        END_IF
    ELSIF tonTotal.Q THEN                      // 事件缺失：超时接管（上界残差回灌断链亦不再挂死）
        _bFail := TRUE;  _uFault := DL_ISR_C_TMO;  _eState := E_DL_IterRunnerPhase.eFail;
    END_IF

E_DL_IterRunnerPhase.eRun:
    IF _bFed THEN
        _bFed := FALSE;  _nIter := _nIter + 1;              // 计数唯一写入点
        IF ((_fFa > 0.0) AND (_fFedF < 0.0)) OR ((_fFa < 0.0) AND (_fFedF > 0.0)) THEN
            _fB := _fFedX;  _fFb := _fFedF;                 // 回灌点与下界异号：替上界
        ELSE
            _fA := _fFedX;  _fFa := _fFedF;
        END_IF
        IF ABS(_fFedF) <= DL_ISR_EPS THEN
            _eState := E_DL_IterRunnerPhase.eDone;          // 残差达标
        ELSIF ABS(_fB - _fA) <= fTol THEN
            _eState := E_DL_IterRunnerPhase.eDone;          // 宽度达标
        ELSIF (nIterMax > 0) AND (_nIter >= nIterMax) THEN
            _bFail := TRUE;  _uFault := DL_ISR_C_ITER;
            _eState := E_DL_IterRunnerPhase.eFail;
        ELSE
            _fXCur := NextTrial(nSel := nMethod, fA := _fA, fB := _fB, fFa := _fFa,
                                fFb := _fFb, fXPrev := _fFedX, fFxPrev := _fFedF);
        END_IF
    ELSIF tonTotal.Q THEN                      // 事件缺失：超时接管（R275 事件优先）
        _bFail := TRUE;  _uFault := DL_ISR_C_TMO;  _eState := E_DL_IterRunnerPhase.eFail;
    END_IF

E_DL_IterRunnerPhase.eDone:
    IF rtStart.Q THEN                          // 启动沿重开一轮
        _bFed := FALSE;  _nIter := 0;  _fA := fXLo;  _fB := fXHi;  _fXCur := fXLo;
        _eState := E_DL_IterRunnerPhase.eEvalLo;
    END_IF

E_DL_IterRunnerPhase.eFail:
    _bFail := TRUE;                            // 失败相驻留：码位锁存回放

E_DL_IterRunnerPhase.eFault:
    _bFault := TRUE;                           // 故障相驻留：出口保持安全值

ELSE
    _bFault := TRUE;  _uFault := DL_ISR_C_ILL;  _eState := E_DL_IterRunnerPhase.eFault;
END_CASE

(* 段 5：故障迁相闸（置于解除段之后，R274） *)
IF _bFault AND (_eState <> E_DL_IterRunnerPhase.eFault) THEN
    _eState := E_DL_IterRunnerPhase.eFault;
END_IF

(* 段 6：统一出口段（判据位与实值单点裁决，N4） *)
bDone := (_eState = E_DL_IterRunnerPhase.eDone);
bError := _bFault OR _bFail;  uErrId := _uFault;  nIterOut := _nIter;
IF (_fXCur <> _fXCur) OR ((_fXCur - _fXCur) <> (_fXCur - _fXCur)) THEN
    fXOut := 0.0;                              // 非有限兜底（N1）
ELSE
    fXOut := _fXCur;
END_IF
IF (_fFedF <> _fFedF) OR ((_fFedF - _fFedF) <> (_fFedF - _fFedF)) THEN
    fResid := 0.0;
ELSE
    fResid := _fFedF;
END_IF
END_FUNCTION_BLOCK

(* ---- FB_DL_KalmanFilter1D.st ---- *)
(*==============================================================================
 * 组件名称 (Component)  : FB_DL_KalmanFilter1D
 * 所属子库 (Sublibrary) : DL_Algo
 * 当前版本 (Version)    : 1.0.0
 * 兼容性   (Platform)   : CODESYS 3.5+ / TwinCAT 3 / 汇川 InoProShop / 施耐德 Machine Expert
 *                         仅依赖 Standard.library（TON / R_TRIG / ABS），零厂商私有库
 * 功能描述 (Function)   : 标量卡尔曼滤波。状态 _fX 与协方差 _fP，逐拍「预测 → 更新」两段：
 *                         预测 _fP := _fP + fQ（随机游走过程噪声）；更新按标量卡尔曼增益
 *                         K = _fP / (_fP + fR)，用新息 |fMeas - _fX| 修正状态并压缩协方差。
 *                         野值门限：新息绝对值超 fInnovLimit → 本拍拒收（bRejected = TRUE，
 *                         不更新状态，协方差保留预测后的增大值，使下一拍更容易接受真变化）。
 *                         协方差发散保护：_fP > fPMax 持续 tDivTime → 用当拍实测重初始化并
 *                         置信息级。失能 bEnable = FALSE → 直通 fMeas 并**冻结协方差**（不归零，
 *                         保证恢复使能时无扰）。
 * 接口     (Interface)  : 输入 fMeas 实测值、fQ 过程噪声、fR 测量噪声、fInnovLimit 新息门限、
 *                         fPMax 协方差发散上限、tDivTime 发散确认时间、bEnable 使能、bReset 复位；
 *                         输出 fOut 滤波值、fPOut 当前协方差、bRejected 本拍拒收单拍位、
 *                         bDiverged 本拍重初始化单拍位、eState / eCause / bError / nErrId。
 * 边界     (Boundary)   : ① 组态闸：fQ / fR / fInnovLimit / fPMax 任一 <= 0.0、tDivTime <= T#0S、
 *                         或任一浮点引脚为 NaN → 故障锁存（NaN 自反判为判等禁令唯一例外）；
 *                         ② 除法前判除子：_fP + fR <= DL_FLOAT_EPS 时跳过更新（不产生 Inf）；
 *                         ③ 新息与状态全走容差比较，禁 `=` / `<>` 判量值；
 *                         ④ NaN 实测 → 本拍整体拒收并置信息级，**不让 NaN 进入 _fP / _fX**
 *                         （R133 / R135：非有限值绝不写入保持槽）；
 *                         ⑤ TON 一枚 + R_TRIG 一枚段 0 无条件周期刷新；
 *                         ⑥ 故障相迁出唯一路径 = bReset 上升沿；⑦ 零全局耦合（无 GVL / 无物理地址）。
 * 输出语义 (Fallback)   : 【R191 声明】bEnable = FALSE → 输出**直通** fMeas（非冻结），协方差冻结
 *                         保持末值；eFault 相 → 输出**冻结保持**末次有效估计（不清零，避免下游
 *                         把 0 当成真测量），bError 同时为真。两分支语义互不相同，均在此显式声明。
 * 解除式   (Release)    : bReset 上升沿 ∧ 组态合法 ∧〔非发散态 ∨ 本次复位已完成协方差重装〕。
 *                         自证可满足（终审两式 1）：复位沿本身在发散态执行 _fP := fR 重装，
 *                         括内第二项即为真，故解除式不存在恒假因子。反例说明：若写成单纯
 *                         「∧ 非发散态」，故障相内 _fP 不再更新 → 该项恒假 → 故障永久不可恢复，
 *                         属 R152 恒假组合反例，故本件按括内析取式实现。
 * 码表     (Codes)      : 16#0002_03AF 故障级：卡尔曼滤波故障总码（组态非法 / 非法相位），
 *                         锁存至 bReset 上升沿，归因由 eCause 承载（R190 单件单总码）；
 *                         16#0002_04B2 信息级：非故障台账事件（野值拒收 / 发散重初始化 / 除子退化跳过）。
 *                         加码反证（R90）：三类信息事件均不改变 eCause 与 bError，且 fOut 仍为
 *                         可用值，故须留痕；三类共用一码的依据是「都只要求留痕、不要求区分动作」，
 *                         区分由 bRejected / bDiverged 两个专用布尔出口承担，无需第二个码位。
 *                         码段说明：0002 段故障子带 03xx / 信息子带 04xx，本件取 03AF / 04B2
 *                         （源码实扫该两槽为空，续接同子带已用最大值，未回填碎片孔洞）。
 * 开源溯源 (Origin)     : 道莅自研 clean-room（参考公开标量卡尔曼递推式与参数域，零代码行复制）
 * 修订历史 (Revision)   : 2026-11-19  v1.0.0  R45 首版（批次 1 · 序号 5）
 *==============================================================================*)

TYPE E_DL_Kf1State :
(
    eIdle  := 0,     // 失能待使能（直通输出） / Idle, disabled, pass-through output
    eRun   := 10,    // 滤波运行 / Filtering in run
    eFault := 90     // 故障锁存相 / Fault latched phase
);
END_TYPE

TYPE E_DL_Kf1Cause :
(
    eNone       := 0,   // 无故障成因 / No cause
    eCfgIllegal := 1,   // 组态非法（含 NaN 参数） / Illegal configuration, including NaN parameters
    ePhaseBad   := 2    // 非法相位兜底 / Illegal phase fallback
);
END_TYPE

FUNCTION_BLOCK FB_DL_KalmanFilter1D
VAR_INPUT
    fMeas       : REAL := 0.0;          // 实测值 [工程单位] / Measured value
    fQ          : REAL := 0.01;         // 过程噪声方差，域 > 0.0 [工程单位²] / Process noise variance, domain > 0.0
    fR          : REAL := 0.10;         // 测量噪声方差，域 > 0.0 [工程单位²] / Measurement noise variance, domain > 0.0
    fInnovLimit : REAL := 5.0;          // 新息门限（野值判据），域 > 0.0 [工程单位] / Innovation limit, domain > 0.0
    fPMax       : REAL := 100.0;        // 协方差发散上限，域 > 0.0 [工程单位²] / Covariance divergence limit, domain > 0.0
    tDivTime    : TIME := T#5S;         // 发散确认时间，域 > T#0S [ms] / Divergence confirm time, domain > T#0S
    bEnable     : BOOL := TRUE;         // 滤波使能，FALSE 时直通并冻结协方差 [-] / Enable, FALSE passes through and freezes covariance
    bReset      : BOOL := FALSE;        // 复位命令，上升沿清故障 [-] / Reset command, rising edge clears fault
END_VAR
VAR_OUTPUT
    fOut        : REAL;                 // 滤波输出值（故障相冻结保持末值） [工程单位] / Filtered output, frozen in fault
    fPOut       : REAL;                 // 当前协方差 [工程单位²] / Current covariance
    bRejected   : BOOL;                 // 本拍野值拒收单拍位 [-] / Single-scan outlier rejection flag
    bDiverged   : BOOL;                 // 本拍发散重初始化单拍位 [-] / Single-scan divergence reinit flag
    eState      : E_DL_Kf1State;        // 状态出口，段 6 单点映射 / State outlet
    eCause      : E_DL_Kf1Cause;        // 故障成因出口（R190 归因唯一） / Fault cause outlet
    bError      : BOOL;                 // 故障锁存标志 [-] / Fault latch flag
    nErrId      : UDINT;                // 事件码，0 = 无事件 / Event code, 0 = no event
END_VAR
VAR
    _eState     : E_DL_Kf1State := E_DL_Kf1State.eIdle;   // 内部相位（CASE 唯一写入目标） / Internal phase
    _eCause     : E_DL_Kf1Cause := E_DL_Kf1Cause.eNone;   // 故障成因锁存（锁存量） / Latched cause
    tonDiv      : TON;                  // 发散确认计时，段 0 无条件调用 / Divergence confirm timer
    rtReset     : R_TRIG;               // 复位沿实例，段 0 无条件调用 / Reset edge
    _fX         : REAL;                 // 状态估计（锁存量） [工程单位] / State estimate, latched
    _fP         : REAL;                 // 状态协方差（锁存量） [工程单位²] / State covariance, latched
    _fInnov     : REAL;                 // 本拍新息 [工程单位] / Innovation this scan
    _fK         : REAL;                 // 本拍卡尔曼增益 [-] / Kalman gain this scan
    _fDen       : REAL;                 // 更新除子 _fP + fR [工程单位²] / Update divisor _fP + fR
    _bInit      : BOOL;                 // 首次初始化完成位（锁存量） [-] / Initialized flag, latched
    _bNonFin    : BOOL;                 // 实测非有限当拍量 [-] / Non-finite measurement this scan
    _bDivCond   : BOOL;                 // 协方差超上限当拍量 [-] / Covariance above limit this scan
    _bCfgBad    : BOOL;                 // 组态非法当拍量 [-] / Illegal configuration
    _bReinit    : BOOL;                 // 本次复位已做协方差重装当拍量 [-] / Covariance re-armed by this reset
    _bFault     : BOOL;                 // 故障锁存位（锁存量） / Latched fault bit
    _uFault     : UDINT;                // 故障码锁存（锁存量） / Latched fault code
    _uInfo      : UDINT;                // 信息码，每拍重算 / Info code, recomputed each scan
END_VAR
VAR CONSTANT
    DL_FLOAT_EPS : REAL := 1.0E-6;      // 浮点判零容差（除子与判等统一口径） [工程单位²] / Float epsilon for zero tests [unit2]
END_VAR

(* —— 段 0：当拍判据派生 + 定时器与沿实例无条件周期刷新 —— *)
_bNonFin := (fMeas <> fMeas) OR ((fMeas - fMeas) <> (fMeas - fMeas));       // 实测 NaN 自反 + Inf 差值自减双判（判等禁令唯一例外） / NaN and Inf detection
_bDivCond := _fP > fPMax;                                                   // 协方差超上限当拍量 / Covariance above limit
_bCfgBad := (fQ <> fQ) OR (fR <> fR) OR (fInnovLimit <> fInnovLimit) OR (fPMax <> fPMax)   // 参数 NaN 组态闸（R151 覆盖每个引脚） / NaN config gate covering every pin
            OR (fQ <= 0.0) OR (fR <= 0.0) OR (fInnovLimit <= 0.0) OR (fPMax <= 0.0)        // 正域组态闸 / Positive-domain config gate
            OR (tDivTime <= T#0S);                                                          // 时间组态闸 / Time config gate
rtReset(CLK := bReset);                                                     // 复位沿，每拍必调（R228A） / Reset edge, called every scan
tonDiv(IN := _bDivCond AND bEnable, PT := tDivTime);                        // 发散确认计时，IN 由判据派生 / Divergence timer, IN derived from verdict

(* —— 段 1：单拍量预清零（锁存量与实例不入清单，R107） —— *)
_uInfo     := 16#0000_0000;        // 信息码每拍重算 / Info recomputed every scan
bRejected  := FALSE;               // 拒收位每拍预清，唯一分支置位（R44 单拍脉冲范式） / Reject flag preset, set in one branch only
bDiverged  := FALSE;               // 重初始化位每拍预清 / Divergence flag preset
_bReinit   := FALSE;               // 复位重装标记每拍预清 / Reset re-arm marker preset
nErrId     := 16#0000_0000;        // 事件码缺省无事件 / Event code default none
bError     := FALSE;               // 故障标志每拍预清，故障分支同拍置位（R45 配对） / Flag preset

(* —— 段 2：复位沿（含发散重装）+ 组态域闸 —— *)
IF rtReset.Q THEN                                                        // 当拍复位沿 / current-scan reset edge
    _bFault := FALSE;                                                    // 清故障锁存位（锁存量） / Clear fault latch
    _uFault := 16#0000_0000;                                             // 清故障锁存码（锁存量） / Clear latched code
    _eCause := E_DL_Kf1Cause.eNone;                                      // 清成因（锁存量） / Clear latched cause
    IF _bDivCond AND (NOT _bNonFin) THEN                                 // 发散态复位：协方差重装（解除可达性关键） / Divergent reset re-arms covariance
        _fP := fR;                                                       // 协方差按测量噪声重装 / Covariance re-armed to measurement noise
        _fX := fMeas;                                                    // 状态按当拍实测重装 / State re-armed to current measurement
        _bReinit := TRUE;                                                // 标记本次复位已完成重装 / Mark re-arm done by this reset
    END_IF
    IF _eState = E_DL_Kf1State.eFault THEN
        _eState := E_DL_Kf1State.eIdle;                                  // 故障相迁出唯一路径 / Sole exit from fault phase
    END_IF
END_IF
IF _bCfgBad THEN                                                         // 组态域闸 / Configuration gate
    _uFault := 16#0002_03AF;                                             // 故障级：卡尔曼滤波故障总码 / Fault-level: filter fault code
    _bFault := TRUE;
    bError  := TRUE;                                                     // 故障标志同拍置位（R45 配对） / Error flag set same scan
    _eCause := E_DL_Kf1Cause.eCfgIllegal;                                // 归因：组态非法 / Cause: illegal configuration
END_IF

(* —— 段 3：首次初始化（仅在无故障且实测有限时取首值） —— *)
IF (NOT _bFault) AND (NOT _bInit) AND (NOT _bNonFin) THEN
    _fX := fMeas;                                                        // 首值取实测 / First value from measurement
    _fP := fR;                                                           // 协方差取测量噪声 / Covariance from measurement noise
    _bInit := TRUE;                                                      // 初始化完成（锁存量） / Initialization done
END_IF

(* —— 段 4：预测 → 更新（仅运行态执行） —— *)
IF (NOT _bFault) AND bEnable AND _bInit AND (NOT _bNonFin) THEN
    _fP := _fP + fQ;                                                     // 预测：协方差增大 / Predict, covariance grows
    IF tonDiv.Q THEN                                                     // 发散确认到：用实测重初始化 / Divergence confirmed, reinit from measurement
        _fX := fMeas;
        _fP := fR;
        bDiverged := TRUE;                                               // 单拍位：本拍做过重初始化 / Single-scan reinit flag
        _uInfo := 16#0002_04B2;                                          // 信息级：发散重初始化留痕 / Info: divergence reinit recorded
    ELSE
        _fInnov := fMeas - _fX;                                          // 新息 / Innovation
        IF ABS(_fInnov) > fInnovLimit THEN                               // 野值门限 / Outlier gate
            bRejected := TRUE;                                           // 单拍位：本拍拒收 / Single-scan reject flag
            _uInfo := 16#0002_04B2;                                      // 信息级：野值拒收留痕 / Info: outlier rejection recorded
        ELSE
            _fDen := _fP + fR;                                           // 更新除子 / Update divisor
            IF _fDen > DL_FLOAT_EPS THEN                                 // 除零前置判 / Divide-by-zero guard
                _fK := _fP / _fDen;                                      // 卡尔曼增益 / Kalman gain
                _fX := _fX + _fK * _fInnov;                              // 状态更新 / State update
                _fP := (1.0 - _fK) * _fP;                                // 协方差压缩 / Covariance shrink
            ELSE
                _uInfo := 16#0002_04B2;                                  // 信息级：除子退化跳过 / Info: degenerate divisor skipped
            END_IF
        END_IF
    END_IF
END_IF
IF (NOT _bFault) AND bEnable AND _bNonFin THEN                           // NaN 实测：本拍拒收留痕 / NaN measurement, reject and record
    bRejected := TRUE;                                                   // 单拍位：本拍拒收 / Single-scan reject flag
    _uInfo := 16#0002_04B2;                                              // 信息级：非有限实测拒收 / Info: non-finite measurement rejected
END_IF

(* —— 段 5：故障解除式（R240 全当拍量；括内析取式自证可满足） —— *)
IF rtReset.Q AND (NOT _bCfgBad) AND ((NOT _bDivCond) OR _bReinit) THEN
    _bFault := FALSE;                                                    // 清故障锁存位（锁存量） / Clear fault latch
    _uFault := 16#0000_0000;                                             // 清故障锁存码（锁存量） / Clear latched code
    _eCause := E_DL_Kf1Cause.eNone;                                      // 清成因（锁存量） / Clear latched cause
END_IF

(* —— 段 5A：故障锁存相位迁移闸 —— *)
IF _bFault AND (_eState <> E_DL_Kf1State.eFault) THEN
    _eState := E_DL_Kf1State.eFault;                                     // 锁存即入故障相 / Latch enters fault phase
END_IF

(* —— 段 6：相位机（ENUM 全成员显式标签 + ELSE 兜底，R128） —— *)
CASE _eState OF

E_DL_Kf1State.eIdle:
    IF bEnable AND _bInit AND (NOT _bFault) THEN                         // 出口 1：使能且已初始化 / Enabled and initialized
        _eState := E_DL_Kf1State.eRun;
    ELSIF _bFault THEN                                                   // 出口 2：故障锁存 / Fault latched
        _eState := E_DL_Kf1State.eFault;
    END_IF

E_DL_Kf1State.eRun:
    IF (NOT bEnable) THEN                                                // 出口 1：失能（前置条件消失，R98） / Disabled, precondition gone
        _eState := E_DL_Kf1State.eIdle;
    ELSIF _bFault THEN                                                   // 出口 2：故障锁存 / Fault latched
        _eState := E_DL_Kf1State.eFault;
    END_IF

E_DL_Kf1State.eFault:
    ;                                                                     // 故障相：仅段 5 复位沿可迁出 / Only the reset edge leaves this phase

ELSE
    _uFault := 16#0002_03AF;                                             // 故障级：非法相位兜底（归并总码） / Illegal-phase fallback
    _bFault := TRUE;
    bError  := TRUE;
    _eCause := E_DL_Kf1Cause.ePhaseBad;                                  // 归因：非法相位 / Cause: illegal phase
    _eState := E_DL_Kf1State.eFault;

END_CASE

(* —— 段 7：出口单点映射（名实同源；锁存码回放；故障相显式钳位） —— *)
IF _bFault THEN
    fOut := _fX;                                                         // 故障相冻结保持末次有效估计（R191 声明） / Frozen hold in fault
ELSIF NOT bEnable THEN
    fOut := fMeas;                                                       // 失能相直通实测（R191 声明） / Pass-through when disabled
ELSE
    fOut := _fX;                                                         // 运行相输出状态估计 / Run-phase state estimate
END_IF
IF (fOut <> fOut) OR ((fOut - fOut) <> (fOut - fOut)) THEN                // 出口非有限复检兜底 / Output non-finite recheck
    fOut := 0.0;                                                         // 非有限即归 0，绝不外溢 / Zero out, never propagate
END_IF
fPOut := _fP;                                                            // 协方差出口（锁存量回放） / Covariance outlet
IF _bFault THEN
    nErrId := _uFault;                                                   // 故障锁存码回放 / Replay latched fault code
ELSE
    nErrId := _uInfo;                                                    // 信息码 / Info code
END_IF
bError := _bFault;                                                       // 故障标志与锁存同源（名实双出口，R191） / Flag from latch
eState := _eState;                                                       // 状态出口 / State outlet
eCause := _eCause;                                                       // 成因出口 / Cause outlet

END_FUNCTION_BLOCK

(* ---- FB_DL_LaminatorPressCtrl.st ---- *)
(*
  FB_DL_LaminatorPressCtrl  —  层压机压力-时间闭环（真空段/加压段分离双目标 + 斜坡限速）/ Laminator pressure-time closed loop
  分类 Category : DL_Algo
  码位 Code     : 16#02_3_88
  段位说明      : 86/87 格由频率/三角波发生件启用，本件启用相邻 88 格（一件一码）
  版本 Version  : 1.0.0
  来源 Source   : t2-2-lbp — ROADMAP 原记 Process 属分层误记，闭环控制律按分层判定归 Algo，本轮改判并留痕
  溯源 Origin   : clean-room 实现，层压压力曲线公开工艺语义借鉴，未复制任何源码行
                  （与 FB_DL_RollCompressForceBalance 分工：那件管力平衡，本件管压力曲线跟随）
  功能 Function : 1) 六相顺控 Idle→Evac→RampPress→Hold→Release→Done，真空段/加压段目标分离；
                  2) 加压目标经 FB_DL_RateLimiter 斜坡限速（fRampRateBarS），斜坡中段由
                  FB_DL_CascadePid 主环（压力）+ 副环（执行器阀位反馈）闭环跟随；
                  3) Hold 相按配方时长 tonHold 驻留，压力越保持窗置信息级码（不静默）；
                  4) Release 相泄压 + 缩回，常压与缩回双确认才进 Done。
  边界 Boundary : ① 真空接口契约：iVac.fPressure 为负压值，深度 = −fPressure（取正深度比较）；
                  ② iActuatorFbPct 为加压执行器阀位反馈 [0..100]%（副环 PV，未接线时副环退化跟随）；
                  ③ R228-A 达标声明：四只定时器均单相独占（IN 为单相等式），跨相迁移拍 IN 必断；
                  ④ 组态域闸覆盖全部参与换算引脚；目标越上限钳制置信息级码；
                  ⑤ R228-B 达标声明：eFault 迁出 = bReset 上升沿（段 4 承载），迁出条件
                  「rtReset.Q」为输入引脚，可满足性自证成立，逐字写于此。
  依赖 Depends  : FB_DL_CascadePid / FB_DL_RateLimiter（实例化，引脚按 registry 实名）；
                  FC_DL_Hysteresis（函数调用，bState 由本件成员持有回传）；
                  I_DL_VacuumGenerator / I_DL_Cylinder（注入，不实例化）
  码表 Error codes（本件格 02_3_88，子码步进 +0x100）:
    16#0002_0188 信息级：周期完成（Done 相）
    16#0002_0288 故障级：组态非法（目标/容差/速率/时长域非法），锁存至复位
    16#0002_0388 故障级：段超时（Evac/Ramp/Release 各相独立计时），锁存至复位
    16#0002_0488 故障级：注入件故障（真空 bFault / 气缸 bFault），锁存至复位
    16#0002_0588 故障级：状态机落 ELSE 兜底（非法相位 ID），锁存至复位
    16#0002_0688 信息级：Hold 相压力越保持窗（等待回落，不置故障）
    16#0002_0788 信息级：压力目标越组态上限，已钳制

  修订历史 Revision :
    2026-11-19  v1.0.0  R39 首版（批次 2 · 序号 6）
*)

TYPE E_DL_LamPressState :
(
    eIdle      := 0,    // 空闲：等启动指令 / Idle, waiting for start
    eEvac      := 10,   // 真空段：抽气至真空目标 / Evacuation to vacuum target
    eRampPress := 20,   // 加压段：斜坡升压 + 串级闭环跟随 / Ramp press with cascade loop
    eHold      := 30,   // 保持段：配方时长驻留 + 保持窗监视 / Recipe hold with window watch
    eRelease   := 40,   // 泄压段：放气 + 缩回双确认 / Release, blow-off and retract confirm
    eDone      := 50,   // 完成：周期落定 / Done
    eFault     := 90    // 故障：组态/超时/注入件锁定 / Fault, latched
);
END_TYPE

FUNCTION_BLOCK FB_DL_LaminatorPressCtrl
VAR_INPUT
    bStart          : BOOL := FALSE;      // 启动指令（上升沿）/ Start command
    fVacTargetKpa   : REAL := 85.0;       // 真空段目标深度 [kPa]，域 > 0 / Vacuum segment target depth
    fPressTargetBar : REAL := 1.5;        // 加压段目标压力 [bar]，域 (0, fPressMaxBar] / Press segment target
    fPressMaxBar    : REAL := 2.0;        // 加压组态上限 [bar]，域 > 0 / Press configuration ceiling
    fPressActBar    : REAL := 0.0;        // 压力变送实测 [bar]（主环 PV）/ Measured pressure, master PV
    fActuatorFbPct  : REAL := 0.0;        // 执行器阀位反馈 [%]（副环 PV）/ Actuator position feedback, slave PV
    fPressTolBar    : REAL := 0.05;       // 压力跟随容差 [bar]，域 > 0 / Pressure tracking tolerance
    fRampRateBarS   : REAL := 0.05;       // 加压斜坡速率 [bar/s]，域 > 0 / Press ramp rate
    fKpM            : REAL := 1.0;        // 主环比例增益 [1] / Master loop proportional gain
    tTiM            : TIME := T#5S;       // 主环积分时间 [s] / Master loop integral time
    fKpS            : REAL := 2.0;        // 副环比例增益 [1] / Slave loop proportional gain
    tTiS            : TIME := T#1S;       // 副环积分时间 [s] / Slave loop integral time
    tEvacDur        : TIME := T#60S;      // 真空段配方时长 [ms] / Evacuation recipe duration
    tEvacTimeout    : TIME := T#120S;     // 真空段超时 [ms]，域 > 0 / Evacuation timeout
    tPressTimeout   : TIME := T#180S;     // 加压段超时 [ms]，域 > 0 / Ramp press timeout
    tHoldDur        : TIME := T#120S;     // 保持段配方时长 [ms] / Hold recipe duration
    tReleaseTimeout : TIME := T#60S;      // 泄压段超时 [ms]，域 > 0 / Release timeout
    fAtmVacKpa      : REAL := 2.0;        // 常压确认阈值 [kPa]，域 >= 0 / Atmospheric confirmation threshold
    bReset          : BOOL := FALSE;      // 复位（eFault 迁出唯一沿）/ Reset, sole fault exit edge
END_VAR
VAR_OUTPUT
    fPressSpRamp    : REAL;               // 斜坡限速后的压力设定 [bar] / Rate-limited pressure setpoint
    fPressCmdPct    : REAL;               // 串级闭环输出 [%] / Cascade closed-loop output in percent
    nSegment        : INT;                // 当前段号 [0..3]（0=真空 1=加压 2=保持 3=泄压）/ Segment index
    bCycleDone      : BOOL;               // 周期完成 / Cycle done
    nErrId          : UDINT;              // 事件码，0 = 无事件 / Event code
    eState          : E_DL_LamPressState; // 状态出口，段尾单点映射 / State outlet
END_VAR
VAR_IN_OUT
    iVac      : I_DL_VacuumGenerator;     // 真空发生器引用（注入，不实例化）/ Vacuum generator reference
    iPressCyl : I_DL_Cylinder;            // 压合气缸引用（注入，不实例化）/ Press cylinder reference
END_VAR
VAR
    fbRate     : FB_DL_RateLimiter;       // 斜坡限速实例 / Ramp rate limiter instance
    fbPid      : FB_DL_CascadePid;        // 压力串级闭环实例 / Pressure cascade loop instance
    tonEvacTo  : TON;                     // 真空段超时（单相独占）/ Evacuation timeout, single phase
    tonPressTo : TON;                     // 加压段超时（单相独占）/ Ramp press timeout, single phase
    tonHold    : TON;                     // 保持段配方计时（单相独占，PT 接配方时长）/ Hold recipe timer, single phase
    tonRelTo   : TON;                     // 泄压段超时（单相独占）/ Release timeout, single phase
    tonWch     : TON;                     // 故障观察窗，自复位 / Fault watch window, self-resetting
    rtStart    : R_TRIG;                  // 启动上升沿 / Start rising edge
    rtReset    : R_TRIG;                  // 复位上升沿 / Reset rising edge
    _eState    : E_DL_LamPressState := E_DL_LamPressState.eIdle;  // 内部相位（CASE 唯一写入目标）/ Internal phase
    _rVacDepth : REAL;                    // 真空深度暂存 [kPa] / Vacuum depth scratch
    _rPressTgt : REAL;                    // 钳制后压力目标 [bar] / Clamped press target
    _rSpRamp   : REAL;                    // 斜坡设定中间量 [bar] / Ramped setpoint working value
    _rCmdPct   : REAL;                    // 闭环输出中间量 [%] / Closed-loop output working value
    _bVacOk    : BOOL;                    // 真空到位标志 / Vacuum reached flag
    _bPressOk  : BOOL;                    // 压力入窗标志 / Pressure in-window flag
    _uFault    : UDINT;                   // 故障码锁存 / Latched fault code
    _uInfo     : UDINT;                   // 信息码，每拍重算 / Info code
    _bFault    : BOOL;                    // 故障锁存位 / Latched fault bit
    _bCfgBad   : BOOL;                    // 组态非法聚合 / Configuration invalid aggregate
END_VAR
VAR CONSTANT
    DL_LP_WATCH_PT : TIME := T#2S;      // 故障观察窗 [ms]，自复位 / Fault watch window
    DL_LP_INF_CAP  : REAL := 1.0E15;    // 非有限值筛查幅值上限 / Non-finite screening cap
END_VAR

(* —— 段 0：定时器与边沿无条件周期刷新（R182：调用语句不得置于 IF/CASE 内） —— *)
(* Stage 0, unconditional refresh of timers and edges *)
rtStart(CLK := bStart);                                           // 启动上升沿，每拍必调
rtReset(CLK := bReset);                                           // 复位上升沿，每拍必调
tonWch(IN := (NOT tonWch.Q), PT := DL_LP_WATCH_PT);               // 观察窗自复位（表达式入参）
tonEvacTo(IN := (_eState = E_DL_LamPressState.eEvac), PT := tEvacTimeout);          // 真空段超时（单相独占）
tonPressTo(IN := (_eState = E_DL_LamPressState.eRampPress), PT := tPressTimeout);   // 加压段超时（单相独占）
tonHold(IN := (_eState = E_DL_LamPressState.eHold), PT := tHoldDur);                // 保持配方计时（单相独占，PT=配方时长）
tonRelTo(IN := (_eState = E_DL_LamPressState.eRelease), PT := tReleaseTimeout);     // 泄压段超时（单相独占）

(* —— 段 1：斜坡与串级实例无条件周期刷新（依赖件每拍必调） —— *)
(* Stage 1, dependency instances refreshed unconditionally *)
fbRate(bEnable := TRUE,                                   // 限速器恒使能，跨相平滑（斜坡连续性）
       fIn := _rPressTgt,                                 // 限速输入 = 钳制后目标
       fRateUp := MAX(fRampRateBarS, 1.0E-6),             // 上升速率（下限防零速率卡死）
       fRateDown := MAX(fRampRateBarS, 1.0E-6),           // 下降速率同源
       bTrack := (_eState <> E_DL_LamPressState.eRampPress),   // 非加压相跟踪实测压力（无扰）
       fTrackValue := fPressActBar,                       // 跟踪值 = 实测压力
       tSampleTime := T#100MS);                           // 采样周期口径与限速件默认一致
_rSpRamp := fbRate.fOut;                                  // 斜坡设定中间量
fbPid(bEnable := (_eState = E_DL_LamPressState.eRampPress) OR (_eState = E_DL_LamPressState.eHold),
      fSpMaster := _rSpRamp,                              // 主环设定 = 斜坡设定
      fPvMaster := fPressActBar,                          // 主环 PV = 压力实测
      fPvSlave := fActuatorFbPct,                         // 副环 PV = 阀位反馈
      fKpM := fKpM, tTiM := tTiM, tTdM := T#0S,           // 主环参数（微分关）
      fKpS := fKpS, tTiS := tTiS, tTdS := T#0S,           // 副环参数（微分关）
      rSpSlaveMin := 0.0, rSpSlaveMax := 100.0,           // 副设定域（阀位百分比）
      rOutMin := 0.0, rOutMax := 100.0,                   // 副环输出域
      tSampleTime := T#100MS, bReset := FALSE);           // 采样周期；PID 自身不复位（相切换靠使能门控）
_rCmdPct := fbPid.fOut;                                   // 闭环输出中间量

(* —— 段 2：单拍量预清零（锁存量 _uFault/_bFault 不入清单，R187①） —— *)
_uInfo := 16#0000_0000;             // 信息码每拍重算
bCycleDone := FALSE;                // 完成出口缺省 FALSE（Done 相单点置位）
_bCfgBad := FALSE;                  // 组态非法预清零
nErrId := 16#0000_0000;             // 事件码缺省无事件

(* —— 段 3：组态域闸（覆盖全部参与判据换算的引脚，R151） —— *)
IF (fVacTargetKpa <> fVacTargetKpa) OR (fVacTargetKpa <= 0.0) OR (ABS(fVacTargetKpa) > DL_LP_INF_CAP)
   OR (fPressActBar <> fPressActBar) OR (ABS(fPressActBar) > DL_LP_INF_CAP) THEN
    _bCfgBad := TRUE;               // 真空目标/压力实测非法
END_IF
IF (fPressMaxBar <= 0.0) OR (fPressTolBar <= 0.0) OR (fRampRateBarS <= 0.0) OR (fAtmVacKpa < 0.0) THEN
    _bCfgBad := TRUE;               // 上限/容差/速率/常压阈非法
END_IF
IF (TIME_TO_DINT(tEvacTimeout) <= 0) OR (TIME_TO_DINT(tPressTimeout) <= 0)
   OR (TIME_TO_DINT(tHoldDur) <= 0) OR (TIME_TO_DINT(tReleaseTimeout) <= 0) THEN
    _bCfgBad := TRUE;               // 各段时长/超时非法
END_IF

(* —— 段 4：eFault 迁出沿（R228-B：迁出条件 rtReset.Q 为输入引脚，恒可达） —— *)
IF rtReset.Q THEN
    _bFault := FALSE;               // 清故障锁存位
    _uFault := 16#0000_0000;
    IF _eState = E_DL_LamPressState.eFault THEN
        _eState := E_DL_LamPressState.eIdle;    // 故障相迁出：回空闲（迁出边唯一且可达）
    END_IF
END_IF

(* —— 段 5：过程量只读采集与判据 —— *)
_rVacDepth := -iVac.fPressure;                // 真空深度 = 负压反馈取反 [kPa]（接口契约：负值=真空）
_bVacOk := _rVacDepth >= fVacTargetKpa;       // 真空到位判据（每拍重算）
_bPressOk := ABS(fPressActBar - _rSpRamp) <= fPressTolBar;   // 压力入窗判据（相对斜坡设定）

(* —— 段 6：相位机（只做迁移与单发命令；出口在段 8） —— *)
CASE _eState OF

E_DL_LamPressState.eIdle:
    IF _bCfgBad AND rtStart.Q THEN
        _uFault := 16#0002_0288;            // 故障级：组态非法
        _bFault := TRUE;
        _eState := E_DL_LamPressState.eFault;
    ELSIF rtStart.Q AND (NOT _bCfgBad) THEN
        IF fPressTargetBar > fPressMaxBar THEN
            _rPressTgt := fPressMaxBar;     // 压力目标越上限钳制
            _uInfo := 16#0002_0788;         // 信息级：已钳制
        ELSE
            _rPressTgt := fPressTargetBar;  // 域内直通
        END_IF
        iVac.CmdEvacuate();                 // 单发抽气指令
        _eState := E_DL_LamPressState.eEvac;    // 进真空段
    END_IF

E_DL_LamPressState.eEvac:
    IF (iVac.bFault OR iPressCyl.bFault) THEN
        _uFault := 16#0002_0488;            // 故障级：注入件故障
        _bFault := TRUE;
        iVac.CmdStop();                     // 安全侧全停
        _eState := E_DL_LamPressState.eFault;
    ELSIF tonEvacTo.Q THEN
        _uFault := 16#0002_0388;            // 故障级：真空段超时
        _bFault := TRUE;
        iVac.CmdStop();
        _eState := E_DL_LamPressState.eFault;
    ELSIF _bVacOk AND tonWch.Q THEN
        _eState := E_DL_LamPressState.eRampPress;   // 真空到位（含观察窗防抖）：进加压段
    END_IF

E_DL_LamPressState.eRampPress:
    IF (iVac.bFault OR iPressCyl.bFault) THEN
        _uFault := 16#0002_0488;
        _bFault := TRUE;
        iPressCyl.CmdStop();                // 安全侧停缸
        _eState := E_DL_LamPressState.eFault;
    ELSIF tonPressTo.Q THEN
        _uFault := 16#0002_0388;            // 故障级：加压段超时
        _bFault := TRUE;
        iPressCyl.CmdStop();
        _eState := E_DL_LamPressState.eFault;
    ELSE
        IF NOT iPressCyl.bExtended THEN
            iPressCyl.CmdExtend();          // 未到位则持续请求伸出（缸件内单发化去重）
        END_IF
        IF _bPressOk AND iPressCyl.bExtended THEN
            _eState := E_DL_LamPressState.eHold;    // 压力入窗且到位：进保持段
        END_IF
    END_IF

E_DL_LamPressState.eHold:
    IF (iVac.bFault OR iPressCyl.bFault) THEN
        _uFault := 16#0002_0488;
        _bFault := TRUE;
        iPressCyl.CmdStop();
        _eState := E_DL_LamPressState.eFault;
    ELSIF NOT _bPressOk THEN
        _uInfo := 16#0002_0688;             // 信息级：保持窗越限（等待回落，不置故障）
    ELSIF tonHold.Q THEN
        iVac.CmdBlowOff();                  // 单发放气（保持到点）
        iPressCyl.CmdRetract();             // 单发缩回
        _eState := E_DL_LamPressState.eRelease;     // 进泄压段
    END_IF

E_DL_LamPressState.eRelease:
    IF (iVac.bFault OR iPressCyl.bFault) THEN
        _uFault := 16#0002_0488;
        _bFault := TRUE;
        iPressCyl.CmdStop();
        _eState := E_DL_LamPressState.eFault;
    ELSIF tonRelTo.Q THEN
        _uFault := 16#0002_0388;            // 故障级：泄压段超时
        _bFault := TRUE;
        _eState := E_DL_LamPressState.eFault;
    ELSIF (_rVacDepth <= fAtmVacKpa) AND (NOT iPressCyl.bExtended) THEN
        _eState := E_DL_LamPressState.eDone;    // 常压 + 缩回双确认：进完成相
    END_IF

E_DL_LamPressState.eDone:
    bCycleDone := TRUE;                     // 完成出口（Done 相每拍重申）
    _uInfo := 16#0002_0188;                 // 信息级：周期完成
    IF NOT bStart THEN
        _eState := E_DL_LamPressState.eIdle;    // 指令撤销：回空闲
    END_IF

E_DL_LamPressState.eFault:
    ;                                       // 故障相：等复位沿（段 4 承载迁出）

ELSE
    _uFault := 16#0002_0588;                // 故障级：非法相位 ID 兜底
    _bFault := TRUE;
    _eState := E_DL_LamPressState.eFault;   // 强制回故障相

END_CASE

(* —— 段 7：出口单点映射（名实同源；锁存码回放，禁同拍抹除） —— *)
IF _eState = E_DL_LamPressState.eEvac THEN
    nSegment := 0;                          // 段号 0：真空
ELSIF _eState = E_DL_LamPressState.eRampPress THEN
    nSegment := 1;                          // 段号 1：加压
ELSIF _eState = E_DL_LamPressState.eHold THEN
    nSegment := 2;                          // 段号 2：保持
ELSIF _eState = E_DL_LamPressState.eRelease THEN
    nSegment := 3;                          // 段号 3：泄压
ELSE
    nSegment := -1;                         // Idle/Done/Fault：无有效段号
END_IF
fPressSpRamp := _rSpRamp;                   // 斜坡设定镜像
fPressCmdPct := _rCmdPct;                   // 闭环输出镜像
IF _bFault THEN
    nErrId := _uFault;                      // 故障锁存码回放（不在故障相按当下输入重推）
    bCycleDone := FALSE;                    // 故障相完成出口强制 FALSE（安全侧）
ELSE
    nErrId := _uInfo;                       // 信息码
END_IF
eState := _eState;                          // 状态出口单点映射

END_FUNCTION_BLOCK

(* ---- FB_DL_LeadLagCompensator.st ---- *)
(*
    FB_DL_LeadLagCompensator —— 一阶超前滞后相位校正器
    ------------------------------------------------------------------
    分类      : DL_Algo / ControlLaw
    前缀      : FB_DL_
    版本      : 1.0.0
    溯源      : 超前滞后校正 Kc·(1 + T_lead·s)/(1 + T_lag·s) 为公开经典控制判据（公共知识）；
                Tustin 双线性离散化、在线改参保状态、旁路与保持判决、错误分级与码位
                100% 自有；只借「控制器归算法层且各律独立成块」的分类组织，不复制任何
                实现代码；clean-room 重写，未复制任何闭源厂商源码，参考实现仅限 MIT/Apache 许可
    平台      : 纯 IEC 61131-3，CODESYS V3.5+ / TwinCAT 3 / InoProShop 通用
    作者      : 道莅代码库 · PLC编程专家（R19）
    ------------------------------------------------------------------
    功能说明  : 回路振荡但相位裕度不足时给前向通道加相位超前；抑制低频扰动时加滞后。
                离散化用 Tustin：a0 = 2·T_lag/Ts + 1，b0 = Kc·(1 + 2·T_lead/Ts)/a0，
                b1 = Kc·(1 − 2·T_lead/Ts)/a0，a1 = (1 − 2·T_lag/Ts)/a0。
                核心防御：① 采样周期越域或滞后时间小于采样周期，离散化极点会出单位圆，
                   此时故障级 2910 并旁路（宁可直通，不可输出病态波形）；
                ② 归一化分母 a0 前置防零判据，绝不裸除；
                ③ 增益非有限或近零即故障级 2911 并旁路——增益 0 会把回路静默掐死，
                   比报错更危险；
                ④ 输入非有限时输出保持末次有效且不旁路（旁路会把毒值直接注入执行器）；
                ⑤ 在线改参逐项比对并重算系数，历史状态保留不清零，切换无扰；
                ⑥ 输出双侧限幅，超限置 bSaturated。
                职责边界：前馈归 FeedforwardComp，纯滞后补偿归 SmithPredictor，各类滤波另件。
    错误码    : 16#0002_2901 时间常数超域已钳位 / 在线改参已重算系数（状态保留）/ 输出限幅生效——信息级，正常防御
                16#0002_2902 预留禁用（信息级，不得挪用）
                16#0002_2910 采样周期或滞后时间非法（离散化失效），旁路输出——故障级，fOut = fIn
                16#0002_2911 增益非有限或近零、输入非有限——故障级，输出保持末次有效
                16#0002_2912 预留禁用（故障级，不得挪用）
    码位总账  : 16#0002_2901 用 / 16#0002_2902 预留 ｜ 16#0002_2910 用 / 16#0002_2911 用 / 16#0002_2912 预留
    状态机    : R6 标注 N/A —— 本组件为纯函数无顺序状态机，无 CASE 可写，非法状态不可能出现
                （旁路/正常由单比特判决在段内直接给出，不存在顺序态）
    采样约定  : fbTrigReset 在本体首部无条件刷新；差分式为直接 I 型（fX1 / fY1 两状态量），
                与直接 II 型转置（单状态量）数学等价，选 I 型以保留输入输出历史供 HMI
                与改参连续性观测；时间基准全部来自 tSampleTime 引脚。
    修订记录  : 2026-11-16 v1.0.0 首次入库（R19）
*)
FUNCTION_BLOCK FB_DL_LeadLagCompensator
VAR_INPUT
    bEnable         : BOOL;                   // 使能，FALSE 旁路（输出 = 输入）/ enable, FALSE bypasses the block, output equals input
    bReset          : BOOL;                   // 复位，上升沿清内部状态 / reset, rising edge clears the internal state
    fIn             : REAL := 0.0;            // 输入（一般接偏差）[用户单位] / input, usually the control error [user unit]
    fGain           : REAL := 1.0;            // 静态增益 Kc [无量纲]，范围 -1000.0~1000.0，禁 0 / static gain [dimensionless], range -1000.0~1000.0, zero forbidden
    tLeadTime       : TIME := T#100MS;        // 超前时间常数 [ms]，范围 0~60000 / lead time constant [ms], range 0~60000
    tLagTime        : TIME := T#1S;           // 滞后时间常数 [ms]，范围 1~600000，必须 ≥ 采样周期 / lag time constant [ms], range 1~600000, must be >= the sample time
    tSampleTime     : TIME := T#100MS;        // 采样周期 [ms]，范围 1~10000 / sample time [ms], range 1~10000
    fOutLimit       : REAL := 1.0E6;          // 输出幅值限幅 [用户单位]，必须 > 0 / output magnitude limit [user unit], must be > 0
END_VAR
VAR_OUTPUT
    fOut            : REAL;                   // 校正后输出 [用户单位] / compensated output [user unit]
    bBypass         : BOOL;                   // 旁路中（参数非法或未使能）/ bypassed, illegal parameters or disabled
    bSaturated      : BOOL;                   // 输出被限幅 / output clamped
    uCoeffRev       : UDINT;                   // 系数重算次数（在线改参监视）[次] / coefficient recompute count [times]
    eErr            : UDINT;                  // 错误码，0=正常 / error id, 0=ok
    bError          : BOOL;                   // 故障标志，eErr 为故障级时 TRUE / error flag, TRUE on fault-level eErr
END_VAR
VAR
    fbTrigReset     : R_TRIG;                 // 复位上升沿实例，本体首部无条件刷新 / reset edge instance, refreshed unconditionally
    fB0             : REAL;                   // Tustin 归一化前向零次系数 [无量纲] / normalised feedforward zero-order coefficient
    fB1             : REAL;                   // Tustin 归一化前向一次系数 [无量纲] / normalised feedforward first-order coefficient
    fA1             : REAL;                   // Tustin 归一化反馈一次系数 [无量纲] / normalised feedback first-order coefficient
    fA0             : REAL;                   // Tustin 归一化分母（防零判据对象）[无量纲] / normalisation denominator, the zero guard target
    fX1             : REAL;                   // 上一拍输入历史 [用户单位] / previous input history [user unit]
    fY1             : REAL;                   // 上一拍输出历史 [用户单位] / previous output history [user unit]
    fPrevK          : REAL;                   // 上一拍增益，改参检测用 [无量纲] / previous gain for change detection [dimensionless]
    fPrevTl         : REAL;                   // 上一拍超前时间，改参检测用 [s] / previous lead time for change detection [s]
    fPrevTg         : REAL;                   // 上一拍滞后时间，改参检测用 [s] / previous lag time for change detection [s]
    fPrevTs         : REAL;                   // 上一拍采样周期，改参检测用 [s] / previous sample time for change detection [s]
    tLeadSec        : REAL;                   // 超前时间常数的秒值 [s] / lead time constant in seconds [s]
    tLagSec         : REAL;                   // 滞后时间常数的秒值 [s] / lag time constant in seconds [s]
    tTsSec          : REAL;                   // 采样周期的秒值 [s] / sample time in seconds [s]
    fLeadEff        : REAL;                   // 钳位后的超前时间 [s] / clamped lead time [s]
    fLagEff         : REAL;                   // 钳位后的滞后时间 [s] / clamped lag time [s]
    fLimitEff       : REAL;                   // 钳位后的输出限幅 [用户单位] / clamped output limit [user unit]
    bParamChg       : BOOL;                   // 在线改参标志 / parameter change flag
    bInit           : BOOL := FALSE;          // 首扫标志，初值 FALSE，判据 NOT bInit / first-scan flag, initial FALSE, tested with NOT
    nDtMs           : DINT;                   // 采样周期毫秒整数 [ms] / sample time in integer milliseconds [ms]
END_VAR
VAR CONSTANT
    DL_LL_LEAD_MAX   : TIME := T#60S;         // 超前时间上限 [ms] / lead time upper bound [ms]
    DL_LL_LAG_MAX    : TIME := T#600S;        // 滞后时间上限 [ms] / lag time upper bound [ms]
    DL_LL_GAIN_MAX   : REAL := 1000.0;        // 增益绝对值上限 [无量纲] / gain magnitude upper bound [dimensionless]
    DL_LL_DT_MAX     : TIME := T#10S;         // 采样周期上限 [ms] / sample time upper bound [ms]
    DL_LL_DT_MIN     : TIME := T#1MS;         // 采样周期下限 [ms] / sample time lower bound [ms]
    DL_FLOAT_EPS     : REAL := 1.0E-6;        // 浮点判等容差 [无量纲] / float equality tolerance [dimensionless]
    DL_LL_MICRO      : REAL := 1.0E-6;        // 微秒级容差，离散系数判定用 [无量纲] / micro tolerance for the discrete coefficients
    DL_LL_MS_PER_S   : REAL := 1000.0;        // 毫秒到秒换算因子 [ms/s] / milliseconds per second [ms/s]
    DL_LL_TWO        : REAL := 2.0;           // Tustin 分子常数 2 [无量纲] / Tustin numerator constant two [dimensionless]
    DL_LL_INF_GUARD  : REAL := 1.0E38;        // 非有限幅值判定阈值 [无量纲] / non-finite magnitude guard [dimensionless]
    DL_LL_ONE        : REAL := 1.0;           // 一值常量，归一化式用 [无量纲] / one constant used by the normalisation [dimensionless]
    DL_LL_CNT_MAX    : UDINT := 16#FFFF_FFFE; // 重算计数饱和值 [次] / recompute counter saturation value [times]
    DL_LL_ZERO       : REAL := 0.0;           // 零值常量，避免裸字面量 [无量纲] / zero constant, avoids a bare literal [dimensionless]
END_VAR

// 段 1｜边沿实例无条件周期刷新（红线：严禁放入条件分支）/ segment 1, unconditional edge refresh
fbTrigReset(CLK := bReset);

// 段 2｜输出与状态预置 / segment 2, preset outputs and status
eErr := 0;                                    // 预置无错误 / preset no error
bError := FALSE;                              // 预置无故障 / preset no fault
bBypass := FALSE;                             // 预置非旁路 / preset not bypassed
bSaturated := FALSE;                          // 预置未饱和 / preset not saturated

// 段 3｜首扫初始化（唯一合法范式：初值 FALSE，判据 NOT bInit）/ segment 3, first-scan initialisation
IF NOT bInit THEN
    fX1 := DL_LL_ZERO;                        // 输入历史清零 / clear the input history
    fY1 := DL_LL_ZERO;                        // 输出历史清零 / clear the output history
    fPrevK := DL_LL_GAIN_MAX;                 // 上一拍增益置哨兵值，首拍必触发重算 / sentinel forces a recompute on the first scan
    fPrevTl := -DL_LL_TWO;                    // 相同哨兵策略 / same sentinel strategy
    fPrevTg := -DL_LL_TWO;                    // 相同哨兵策略 / same sentinel strategy
    fPrevTs := -DL_LL_TWO;                    // 相同哨兵策略 / same sentinel strategy
    bInit := TRUE;                            // 首扫只做一次 / first scan runs once only
END_IF

// 段 4｜使能闸：未使能直接旁路 / segment 4, enable gate bypasses the block
IF NOT bEnable THEN
    bBypass := TRUE;                          // 标记旁路 / flag the bypass
    fOut := fIn;                              // 旁路即直通 / bypass means straight through
    RETURN;                                   // 失能即出口 / disabled is the exit
END_IF

// 段 5｜采样周期与滞后时间闸（离散化失效时宁可直通）/ segment 5, discretisation validity gate
IF (tSampleTime < DL_LL_DT_MIN) OR (tSampleTime > DL_LL_DT_MAX) THEN
    eErr := 16#0002_2910;                     // 采样周期非法故障码 / illegal sample time fault id
    bError := TRUE;                           // 置故障标志 / raise the error flag
    bBypass := TRUE;                          // 旁路输出 / bypass the output
    fOut := fIn;                              // 直通，不输出病态波形 / straight through, never emit a pathological waveform
    RETURN;                                   // 故障级提前返回 / early return on fault
END_IF
IF tLagTime < tSampleTime THEN
    eErr := 16#0002_2910;                     // 滞后时间小于采样周期，极点会出单位圆 / a lag shorter than the sample time pushes the pole outside the unit circle
    bError := TRUE;                           // 置故障标志 / raise the error flag
    bBypass := TRUE;                          // 旁路输出 / bypass the output
    fOut := fIn;                              // 直通 / straight through
    RETURN;                                   // 故障级提前返回 / early return on fault
END_IF

// 段 6｜增益闸（增益 0 会把回路静默掐死，必须报错并旁路）/ segment 6, gain gate
IF (fGain <> fGain) OR (fGain > DL_LL_INF_GUARD) OR (fGain < -DL_LL_INF_GUARD)
   OR (ABS(fGain) <= DL_FLOAT_EPS) OR (ABS(fGain) > DL_LL_GAIN_MAX) THEN
    eErr := 16#0002_2911;                     // 增益非法故障码 / illegal gain fault id
    bError := TRUE;                           // 置故障标志 / raise the error flag
    bBypass := TRUE;                          // 旁路输出 / bypass the output
    fOut := fIn;                              // 直通 / straight through
    RETURN;                                   // 故障级提前返回 / early return on fault
END_IF

// 段 7｜时间常数域钳位（超上限只钳位并留信息码）/ segment 7, time constant domain clamp
fLeadEff := DINT_TO_REAL(TIME_TO_DINT(tLeadTime)) / DL_LL_MS_PER_S; // 超前时间换算为秒 [s] / lead time in seconds [s]
fLagEff := DINT_TO_REAL(TIME_TO_DINT(tLagTime)) / DL_LL_MS_PER_S;   // 滞后时间换算为秒 [s] / lag time in seconds [s]
nDtMs := TIME_TO_DINT(tSampleTime);           // 采样周期取整数毫秒 [ms] / sample time in integer milliseconds [ms]
tTsSec := DINT_TO_REAL(nDtMs) / DL_LL_MS_PER_S; // 采样周期换算为秒，除子为常量 [s] / sample time in seconds, divisor is a constant [s]
IF fLeadEff < DL_LL_ZERO THEN
    fLeadEff := DL_LL_ZERO;                   // 超前时间为负无物理意义 / a negative lead time has no physical meaning
    eErr := 16#0002_2901;                     // 信息级：已钳位 / info level, clamped
END_IF
IF fLeadEff > (DINT_TO_REAL(TIME_TO_DINT(DL_LL_LEAD_MAX)) / DL_LL_MS_PER_S) THEN
    fLeadEff := DINT_TO_REAL(TIME_TO_DINT(DL_LL_LEAD_MAX)) / DL_LL_MS_PER_S; // 超前时间超上限钳位 [s] / clamp the lead time at its upper bound [s]
    eErr := 16#0002_2901;                     // 信息级：已钳位 / info level, clamped
END_IF
IF fLagEff > (DINT_TO_REAL(TIME_TO_DINT(DL_LL_LAG_MAX)) / DL_LL_MS_PER_S) THEN
    fLagEff := DINT_TO_REAL(TIME_TO_DINT(DL_LL_LAG_MAX)) / DL_LL_MS_PER_S; // 滞后时间超上限钳位 [s] / clamp the lag time at its upper bound [s]
    eErr := 16#0002_2901;                     // 信息级：已钳位 / info level, clamped
END_IF
tLeadSec := fLeadEff;                         // 记录生效超前时间 [s] / record the effective lead time [s]
tLagSec := fLagEff;                           // 记录生效滞后时间 [s] / record the effective lag time [s]

// 段 8｜输出限幅参数域钳位（0 或负值会让输出恒 0）/ segment 8, output limit clamp
fLimitEff := fOutLimit;                       // 取入参副本 / copy the input
IF (fLimitEff <> fLimitEff) OR (fLimitEff < DL_FLOAT_EPS) THEN
    fLimitEff := DL_LL_GAIN_MAX;              // 非法限幅退回常量上限 / fall back to the constant bound
    eErr := 16#0002_2901;                     // 信息级：限幅参数已收敛 / info level, the limit was converged
END_IF

// 段 9｜在线改参检测（逐项比对，命中即重算系数并保留历史状态）/ segment 9, online parameter change detection
bParamChg := (ABS(fGain - fPrevK) > DL_FLOAT_EPS)
          OR (ABS(tLeadSec - fPrevTl) > DL_FLOAT_EPS)
          OR (ABS(tLagSec - fPrevTg) > DL_FLOAT_EPS)
          OR (ABS(tTsSec - fPrevTs) > DL_FLOAT_EPS); // 改参判定 / parameter change detection
IF bParamChg THEN
    fA0 := DL_LL_TWO * tLagSec / tTsSec + DL_LL_ONE; // 归一化分母 a0 = 2·T_lag/Ts + 1 / normalisation denominator
    IF ABS(fA0) <= DL_LL_MICRO THEN
        eErr := 16#0002_2910;                 // 分母近零，离散化不可用（前置防零）/ the denominator is near zero, the discretisation is unusable
        bError := TRUE;                       // 置故障标志 / raise the error flag
        bBypass := TRUE;                      // 旁路输出 / bypass the output
        fOut := fIn;                          // 直通 / straight through
        RETURN;                               // 故障级提前返回，绝不裸除 / early return, never divide blindly
    END_IF
    fB0 := fGain * (DL_LL_TWO * tLeadSec / tTsSec + DL_LL_ONE) / fA0; // 前向零次系数 / feedforward zero-order coefficient
    fB1 := fGain * (DL_LL_ONE - DL_LL_TWO * tLeadSec / tTsSec) / fA0; // 前向一次系数 / feedforward first-order coefficient
    fA1 := (DL_LL_ONE - DL_LL_TWO * tLagSec / tTsSec) / fA0;          // 反馈一次系数 / feedback first-order coefficient
    fPrevK := fGain;                          // 记录本拍增益 / remember the gain
    fPrevTl := tLeadSec;                      // 记录本拍超前时间 / remember the lead time
    fPrevTg := tLagSec;                       // 记录本拍滞后时间 / remember the lag time
    fPrevTs := tTsSec;                        // 记录本拍采样周期 / remember the sample time
    IF uCoeffRev < DL_LL_CNT_MAX THEN
        uCoeffRev := uCoeffRev + 1;           // 重算次数饱和加一 / saturating recompute counter
    END_IF
    IF eErr = 0 THEN
        eErr := 16#0002_2901;                 // 信息级：在线改参已重算系数，状态保留 / info level, coefficients recomputed, state kept
    END_IF
    // 历史状态 fX1 / fY1 不清零：改参瞬间无扰，避免输出台阶冲击执行器 / the history is deliberately kept, so a parameter change causes no step
END_IF

// 段 10｜输入非有限闸：输出保持末次有效，且不旁路（旁路会把毒值注入执行器）/ segment 10, non-finite input gate
IF (fIn <> fIn) OR (fIn > DL_LL_INF_GUARD) OR (fIn < -DL_LL_INF_GUARD) THEN
    eErr := 16#0002_2911;                     // 输入非有限故障码 / non-finite input fault id
    bError := TRUE;                           // 置故障标志 / raise the error flag
    RETURN;                                   // 保持末次 fOut，绝不直通 / hold the last output, never pass the poison value through
END_IF

// 段 11｜复位沿清内部状态（在运算之前生效）/ segment 11, reset clears the internal state
IF fbTrigReset.Q THEN
    fX1 := DL_LL_ZERO;                        // 清输入历史 / clear the input history
    fY1 := DL_LL_ZERO;                        // 清输出历史 / clear the output history
END_IF

// 段 12｜直接 I 型差分式（两状态量，系数已归一化）/ segment 12, direct form I difference equation
fOut := fB0 * fIn + fB1 * fX1 - fA1 * fY1;    // y = b0·x + b1·x1 − a1·y1 [用户单位] / the difference equation [user unit]

// 段 13｜结果非有限复检（此时 fY1 仍是上一拍有效输出，可安全回退）/ segment 13, non-finite recheck before the state shift
IF (fOut <> fOut) OR (fOut > DL_LL_INF_GUARD) OR (fOut < -DL_LL_INF_GUARD) THEN
    eErr := 16#0002_2911;                     // 结果非有限，按输入故障同码处理 / a non-finite result shares the input fault id
    bError := TRUE;                           // 置故障标志 / raise the error flag
    fOut := fY1;                              // 回退到上一拍有效输出（位移尚未发生）/ fall back to the previous valid output, the shift has not happened yet
    RETURN;                                   // 出口 / exit
END_IF
IF fOut > fLimitEff THEN
    fOut := fLimitEff;                        // 正向限幅 / clamp the positive side
    bSaturated := TRUE;                       // 标记饱和 / flag the saturation
    eErr := 16#0002_2901;                     // 信息级：输出限幅生效 / info level, the output limit is active
ELSIF fOut < -fLimitEff THEN
    fOut := -fLimitEff;                       // 负向限幅 / clamp the negative side
    bSaturated := TRUE;                       // 标记饱和 / flag the saturation
    eErr := 16#0002_2901;                     // 同一业务语义复用同一信息码 / the same semantics reuses the same info id
END_IF

// 段 15｜状态位移（顺序不可颠倒：运算与限幅全部结束后才移）/ segment 15, state shift at the very end
fX1 := fIn;                                   // 记录本拍输入 / remember this cycle input
fY1 := fOut;                                  // 记录本拍输出 / remember this cycle output
END_FUNCTION_BLOCK
